// ROLL migration prototype. Compile and verify in TIA V19 before commissioning.
// No absolute M aliases: byte/word reads below preserve S5 overlapping memory.
TYPE "ROLL_TimerState"
VERSION : 0.1
STRUCT
    RemainingMs : LReal;
    BaseMs : Int;
    Mode : Int;
    Previous : Bool;
    Q : Bool;
END_STRUCT;
END_TYPE

TYPE "ROLL_CounterState"
VERSION : 0.1
STRUCT
    Value : Int;
    SetPrevious : Bool;
    UpPrevious : Bool;
    DownPrevious : Bool;
END_STRUCT;
END_TYPE

DATA_BLOCK "ROLL_State"
{ S7_Optimized_Access := 'TRUE' }
VERSION : 0.1
NON_RETAIN
VAR
    M : Array[0..255, 0..7] of Bool;
    S5Timers : Array[0..127] of "ROLL_TimerState";
    S5Counters : Array[0..127] of "ROLL_CounterState";
    CurrentProgram : Int := 1;
END_VAR
BEGIN
    M[0, 4] := TRUE;
END_DATA_BLOCK

DATA_BLOCK "ROLL_IO"
{ S7_Optimized_Access := 'TRUE' }
VERSION : 0.1
NON_RETAIN
VAR
    Input : Array[0..127, 0..7] of Bool;
    Output : Array[0..127, 0..7] of Bool;
    Simulation : Bool := TRUE;
    PhysicalOutputsEnabled : Bool := FALSE;
    PhysicalIoConfigured : Bool := FALSE;
    ConversionFault : Bool;
    FirstCycle : Bool := TRUE;
    RuntimeMemory : LReal;
    ClockMs : LReal;
    HmiElapsedMs : LReal;
    HmiLastHeartbeat : DInt;
END_VAR
BEGIN
END_DATA_BLOCK

// Flat, symbolic WinCC interface; TP900 control binding is a separate build step.
DATA_BLOCK "ROLL_HMI"
{ S7_Optimized_Access := 'TRUE' }
VERSION : 0.1
NON_RETAIN
VAR
    Heartbeat : DInt;
    Connected : Bool;
    ManualFunction : Int := 255;
    GroundHeld : Bool;
    WorkHeld : Bool;
    KeyF : Array[1..16] of Bool;
    SelectedProgram : Int := 1;
    RecipeCommand : Int := 1;
    RecipeRequest : DInt;
    RecipeAck : DInt;
    RecipeError : Int;
    CurrentProgram : Int := 1;
    ParameterRequest : DInt;
    ParameterAck : DInt;
    ParameterDb : Int := 15;
    ParameterIndex : Int;
    ParameterValue : DInt;
    ParameterCurrentValue : DInt;
    ParameterSlotPresent : Bool;
    ParameterError : Int;
    Dwell1Seconds : Int := 360;
    Drain1Seconds : Int := 90;
    Ultrasound1 : Bool := TRUE;
    Dwell2Seconds : Int := 240;
    Drain2Seconds : Int := 60;
    Dwell3Seconds : Int := 300;
    Drain3Seconds : Int := 120;
    Dry4Seconds : Int := 400;
    BasketMotion : Int := 1;
    BathLift : Bool;
    ProcessTimer1Units : Int;
    ProcessTimer2Units : Int;
    StatusM : Array[0..255, 0..7] of Bool;
    LogicalOutputs : Array[16..25, 0..7] of Bool;
END_VAR
BEGIN
END_DATA_BLOCK


DATA_BLOCK "ROLL_DB15"
{ S7_Optimized_Access := 'TRUE' }
VERSION : 0.1
NON_RETAIN
VAR
    DW : Array[0..131] of Word;
END_VAR
BEGIN
    DW[0] := W#16#FFFF;
    DW[1] := W#16#FFFF;
    DW[2] := W#16#FFFF;
    DW[3] := W#16#FFFF;
    DW[4] := W#16#FFFF;
    DW[5] := W#16#FFFF;
    DW[6] := W#16#FFFF;
    DW[7] := W#16#FFFF;
    DW[8] := W#16#FFFF;
    DW[9] := W#16#FFFF;
    DW[10] := W#16#FFFF;
    DW[11] := W#16#FFFF;
    DW[12] := W#16#FFFF;
    DW[13] := W#16#FFFF;
    DW[14] := W#16#FFFF;
    DW[15] := W#16#FFFF;
    DW[16] := W#16#FFFF;
    DW[17] := W#16#3360;
    DW[18] := W#16#FFFF;
    DW[19] := W#16#FFFF;
    DW[20] := W#16#FFFF;
    DW[21] := W#16#FFFF;
    DW[22] := W#16#FFFF;
    DW[23] := W#16#FFFF;
    DW[24] := W#16#1010;
    DW[25] := W#16#1020;
    DW[26] := W#16#FFFF;
    DW[27] := W#16#FFFF;
    DW[28] := W#16#FFFF;
    DW[29] := W#16#FFFF;
    DW[30] := W#16#FFFF;
    DW[31] := W#16#3120;
    DW[32] := W#16#3120;
    DW[33] := W#16#2900;
    DW[34] := W#16#FFFF;
    DW[35] := W#16#FFFF;
    DW[36] := W#16#FFFF;
    DW[37] := W#16#FFFF;
    DW[38] := W#16#FFFF;
    DW[39] := W#16#FFFF;
    DW[40] := W#16#FFFF;
    DW[41] := W#16#FFFF;
    DW[42] := W#16#FFFF;
    DW[43] := W#16#FFFF;
    DW[44] := W#16#FFFF;
    DW[45] := W#16#FFFF;
    DW[46] := W#16#FFFF;
    DW[47] := W#16#FFFF;
    DW[48] := W#16#FFFF;
    DW[49] := W#16#FFFF;
    DW[50] := W#16#FFFF;
    DW[51] := W#16#FFFF;
    DW[52] := W#16#FFFF;
    DW[53] := W#16#2120;
    DW[54] := W#16#2120;
    DW[55] := W#16#1010;
    DW[56] := W#16#2060;
    DW[57] := W#16#FFFF;
    DW[58] := W#16#3180;
    DW[59] := W#16#3180;
    DW[60] := W#16#2060;
    DW[61] := W#16#2600;
    DW[62] := W#16#2600;
    DW[63] := W#16#2010;
    DW[64] := W#16#FFFF;
    DW[65] := W#16#2015;
    DW[66] := W#16#FFFF;
    DW[67] := W#16#1050;
    DW[68] := W#16#FFFF;
    DW[69] := W#16#FFFF;
    DW[70] := W#16#FFFF;
    DW[71] := W#16#FFFF;
    DW[72] := W#16#FFFF;
    DW[73] := W#16#FFFF;
    DW[74] := W#16#FFFF;
    DW[75] := W#16#2600;
    DW[76] := W#16#FFFF;
    DW[77] := W#16#2300;
    DW[78] := W#16#FFFF;
    DW[79] := W#16#FFFF;
    DW[80] := W#16#FFFF;
    DW[81] := W#16#FFFF;
    DW[82] := W#16#FFFF;
    DW[83] := W#16#FFFF;
    DW[84] := W#16#FFFF;
    DW[85] := W#16#2120;
    DW[86] := W#16#FFFF;
    DW[87] := W#16#FFFF;
    DW[88] := W#16#FFFF;
    DW[89] := W#16#FFFF;
    DW[90] := W#16#FFFF;
    DW[91] := W#16#FFFF;
    DW[92] := W#16#FFFF;
    DW[93] := W#16#FFFF;
    DW[94] := W#16#FFFF;
    DW[95] := W#16#FFFF;
    DW[96] := W#16#FFFF;
    DW[97] := W#16#FFFF;
    DW[98] := W#16#FFFF;
    DW[99] := W#16#FFFF;
    DW[100] := W#16#FFFF;
    DW[101] := W#16#FFFF;
    DW[102] := W#16#2300;
    DW[103] := W#16#2300;
    DW[104] := W#16#FFFF;
    DW[105] := W#16#FFFF;
    DW[106] := W#16#2010;
    DW[107] := W#16#2015;
    DW[108] := W#16#FFFF;
    DW[109] := W#16#FFFF;
    DW[110] := W#16#FFFF;
    DW[111] := W#16#FFFF;
    DW[112] := W#16#FFFF;
    DW[113] := W#16#FFFF;
    DW[114] := W#16#FFFF;
    DW[115] := W#16#1050;
    DW[116] := W#16#1050;
    DW[117] := W#16#1050;
    DW[118] := W#16#FFFF;
    DW[119] := W#16#FFFF;
    DW[120] := W#16#FFFF;
    DW[121] := W#16#FFFF;
    DW[122] := W#16#FFFF;
    DW[123] := W#16#FFFF;
    DW[124] := W#16#FFFF;
    DW[125] := W#16#FFFF;
    DW[126] := W#16#FFFF;
    DW[127] := W#16#0038;
    DW[128] := W#16#0011;
    DW[129] := W#16#0011;
    DW[130] := W#16#3360;
    DW[131] := W#16#0000;
END_DATA_BLOCK

DATA_BLOCK "ROLL_DB19"
{ S7_Optimized_Access := 'TRUE' }
VERSION : 0.1
NON_RETAIN
VAR
    DW : Array[0..131] of Word;
END_VAR
BEGIN
    DW[0] := W#16#FFFF;
    DW[1] := W#16#0020;
    DW[2] := W#16#0014;
    DW[3] := W#16#FFFF;
    DW[4] := W#16#FFFF;
    DW[5] := W#16#FFFF;
    DW[6] := W#16#FFFF;
    DW[7] := W#16#FFFF;
    DW[8] := W#16#FFFF;
    DW[9] := W#16#FFFF;
    DW[10] := W#16#FFFF;
    DW[11] := W#16#FFFF;
    DW[12] := W#16#FFFF;
    DW[13] := W#16#FFFF;
    DW[14] := W#16#FFFF;
    DW[15] := W#16#FFFF;
    DW[16] := W#16#FFFF;
    DW[17] := W#16#FFFF;
    DW[18] := W#16#FFFF;
    DW[19] := W#16#FFFF;
    DW[20] := W#16#FFFF;
    DW[21] := W#16#FFFF;
    DW[22] := W#16#FFFF;
    DW[23] := W#16#FFFF;
    DW[24] := W#16#FFFF;
    DW[25] := W#16#FFFF;
    DW[26] := W#16#FFFF;
    DW[27] := W#16#FFFF;
    DW[28] := W#16#FFFF;
    DW[29] := W#16#FFFF;
    DW[30] := W#16#FFFF;
    DW[31] := W#16#FFFF;
    DW[32] := W#16#FFFF;
    DW[33] := W#16#FFFF;
    DW[34] := W#16#FFFF;
    DW[35] := W#16#FFFF;
    DW[36] := W#16#FFFF;
    DW[37] := W#16#FFFF;
    DW[38] := W#16#FFFF;
    DW[39] := W#16#FFFF;
    DW[40] := W#16#FFFF;
    DW[41] := W#16#FFFF;
    DW[42] := W#16#FFFF;
    DW[43] := W#16#FFFF;
    DW[44] := W#16#FFFF;
    DW[45] := W#16#FFFF;
    DW[46] := W#16#FFFF;
    DW[47] := W#16#FFFF;
    DW[48] := W#16#FFFF;
    DW[49] := W#16#FFFF;
    DW[50] := W#16#FFFF;
    DW[51] := W#16#FFFF;
    DW[52] := W#16#FFFF;
    DW[53] := W#16#FFFF;
    DW[54] := W#16#FFFF;
    DW[55] := W#16#FFFF;
    DW[56] := W#16#FFFF;
    DW[57] := W#16#FFFF;
    DW[58] := W#16#FFFF;
    DW[59] := W#16#FFFF;
    DW[60] := W#16#FFFF;
    DW[61] := W#16#FFFF;
    DW[62] := W#16#FFFF;
    DW[63] := W#16#FFFF;
    DW[64] := W#16#FFFF;
    DW[65] := W#16#FFFF;
    DW[66] := W#16#FFFF;
    DW[67] := W#16#FFFF;
    DW[68] := W#16#FFFF;
    DW[69] := W#16#FFFF;
    DW[70] := W#16#FFFF;
    DW[71] := W#16#FFFF;
    DW[72] := W#16#FFFF;
    DW[73] := W#16#FFFF;
    DW[74] := W#16#FFFF;
    DW[75] := W#16#FFFF;
    DW[76] := W#16#FFFF;
    DW[77] := W#16#FFFF;
    DW[78] := W#16#FFFF;
    DW[79] := W#16#FFFF;
    DW[80] := W#16#FFFF;
    DW[81] := W#16#FFFF;
    DW[82] := W#16#FFFF;
    DW[83] := W#16#FFFF;
    DW[84] := W#16#FFFF;
    DW[85] := W#16#FFFF;
    DW[86] := W#16#FFFF;
    DW[87] := W#16#FFFF;
    DW[88] := W#16#FFFF;
    DW[89] := W#16#FFFF;
    DW[90] := W#16#FFFF;
    DW[91] := W#16#FFFF;
    DW[92] := W#16#FFFF;
    DW[93] := W#16#FFFF;
    DW[94] := W#16#FFFF;
    DW[95] := W#16#FFFF;
    DW[96] := W#16#FFFF;
    DW[97] := W#16#FFFF;
    DW[98] := W#16#FFFF;
    DW[99] := W#16#FFFF;
    DW[100] := W#16#FFFF;
    DW[101] := W#16#FFFF;
    DW[102] := W#16#FFFF;
    DW[103] := W#16#FFFF;
    DW[104] := W#16#FFFF;
    DW[105] := W#16#FFFF;
    DW[106] := W#16#FFFF;
    DW[107] := W#16#FFFF;
    DW[108] := W#16#FFFF;
    DW[109] := W#16#FFFF;
    DW[110] := W#16#FFFF;
    DW[111] := W#16#FFFF;
    DW[112] := W#16#FFFF;
    DW[113] := W#16#FFFF;
    DW[114] := W#16#FFFF;
    DW[115] := W#16#FFFF;
    DW[116] := W#16#FFFF;
    DW[117] := W#16#FFFF;
    DW[118] := W#16#FFFF;
    DW[119] := W#16#FFFF;
    DW[120] := W#16#FFFF;
    DW[121] := W#16#FFFF;
    DW[122] := W#16#FFFF;
    DW[123] := W#16#FFFF;
    DW[124] := W#16#FFFF;
    DW[125] := W#16#FFFF;
    DW[126] := W#16#FFFF;
    DW[127] := W#16#FFFF;
    DW[128] := W#16#0001;
    DW[129] := W#16#0001;
    DW[130] := W#16#0020;
    DW[131] := W#16#0000;
END_DATA_BLOCK

DATA_BLOCK "ROLL_Recipe1"
{ S7_Optimized_Access := 'TRUE' }
VERSION : 0.1
NON_RETAIN
VAR
    DW : Array[0..41] of Word;
END_VAR
BEGIN
    DW[5] := W#16#2360;
    DW[9] := W#16#2090;
    DW[13] := W#16#0001;
    DW[17] := W#16#2240;
    DW[21] := W#16#2060;
    DW[25] := W#16#2300;
    DW[29] := W#16#2120;
    DW[33] := W#16#2400;
    DW[37] := W#16#0001;
    DW[41] := W#16#0000;
END_DATA_BLOCK

DATA_BLOCK "ROLL_Recipe2"
{ S7_Optimized_Access := 'TRUE' }
VERSION : 0.1
NON_RETAIN
VAR
    DW : Array[0..41] of Word;
END_VAR
BEGIN
    DW[5] := W#16#2360;
    DW[9] := W#16#2090;
    DW[13] := W#16#0001;
    DW[17] := W#16#2240;
    DW[21] := W#16#2060;
    DW[25] := W#16#2300;
    DW[29] := W#16#2120;
    DW[33] := W#16#2400;
    DW[37] := W#16#0001;
    DW[41] := W#16#0000;
END_DATA_BLOCK

DATA_BLOCK "ROLL_DB205"
{ S7_Optimized_Access := 'TRUE' }
VERSION : 0.1
NON_RETAIN
VAR
    DW : Array[0..41] of Word;
END_VAR
BEGIN
    DW[5] := W#16#2360;
    DW[9] := W#16#2090;
    DW[13] := W#16#0001;
    DW[17] := W#16#2240;
    DW[21] := W#16#2060;
    DW[25] := W#16#2300;
    DW[29] := W#16#2120;
    DW[33] := W#16#2400;
    DW[37] := W#16#0001;
    DW[41] := W#16#0000;
END_DATA_BLOCK

FUNCTION "ROLL_GetM" : Word
{ S7_Optimized_Access := 'TRUE' }
VERSION : 0.1
VAR_INPUT
    FirstByte : Int;
    Width : Int;
END_VAR
VAR_TEMP
    b : Int;
    n : Int;
    bit : Int;
    mask : Word;
    result : Word;
END_VAR
BEGIN
    #result := W#16#0000;
    IF (#FirstByte < 0) OR (#FirstByte > 255) OR ((#Width <> 8) AND (#Width <> 16)) OR ((#Width = 16) AND (#FirstByte > 254)) THEN
        "ROLL_IO".ConversionFault := TRUE;
        #ROLL_GetM := #result;
        RETURN;
    END_IF;
    FOR #n := 0 TO (#Width / 8) - 1 DO
        #b := #FirstByte + #n;
        FOR #bit := 0 TO 7 DO
            #mask := SHL(IN := W#16#0001, N := INT_TO_USINT(#bit + (#Width - 8 - 8 * #n)));
            IF "ROLL_State".M[#b, #bit] THEN #result := #result OR #mask; END_IF;
        END_FOR;
    END_FOR;
    #ROLL_GetM := #result;
END_FUNCTION

FUNCTION "ROLL_SetMWord" : Void
{ S7_Optimized_Access := 'TRUE' }
VERSION : 0.1
VAR_INPUT
    FirstByte : Int;
    Value : Word;
END_VAR
VAR_TEMP
    bit : Int;
END_VAR
BEGIN
    IF (#FirstByte < 0) OR (#FirstByte > 254) THEN
        "ROLL_IO".ConversionFault := TRUE;
        RETURN;
    END_IF;
    FOR #bit := 0 TO 7 DO
        "ROLL_State".M[#FirstByte, #bit] := (#Value AND SHL(IN := W#16#0001, N := INT_TO_USINT(#bit + 8))) <> W#16#0000;
        "ROLL_State".M[#FirstByte + 1, #bit] := (#Value AND SHL(IN := W#16#0001, N := INT_TO_USINT(#bit))) <> W#16#0000;
    END_FOR;
END_FUNCTION

FUNCTION "ROLL_GetDW" : Word
{ S7_Optimized_Access := 'TRUE' }
VERSION : 0.1
VAR_INPUT
    DbNumber : Int;
    Index : Int;
END_VAR
BEGIN
    #ROLL_GetDW := W#16#0000;
    IF (#Index < 0) OR (#Index > 131) THEN
        "ROLL_IO".ConversionFault := TRUE;
        RETURN;
    END_IF;
    CASE #DbNumber OF
        15: #ROLL_GetDW := "ROLL_DB15".DW[#Index];
        19: #ROLL_GetDW := "ROLL_DB19".DW[#Index];
        ELSE "ROLL_IO".ConversionFault := TRUE;
    END_CASE;
END_FUNCTION

FUNCTION "ROLL_DecodeBCD" : Int
{ S7_Optimized_Access := 'TRUE' }
VERSION : 0.1
VAR_INPUT
    Value : Word;
END_VAR
VAR_TEMP
    hundreds : Int;
    tens : Int;
    units : Int;
END_VAR
BEGIN
    #hundreds := WORD_TO_INT(SHR(IN := #Value AND W#16#0F00, N := 8));
    #tens := WORD_TO_INT(SHR(IN := #Value AND W#16#00F0, N := 4));
    #units := WORD_TO_INT(#Value AND W#16#000F);
    IF (#hundreds > 9) OR (#tens > 9) OR (#units > 9) THEN
        "ROLL_IO".ConversionFault := TRUE;
        #ROLL_DecodeBCD := -1;
    ELSE
        #ROLL_DecodeBCD := #hundreds * 100 + #tens * 10 + #units;
    END_IF;
END_FUNCTION

FUNCTION "ROLL_EncodeSeconds" : Word
{ S7_Optimized_Access := 'TRUE' }
VERSION : 0.1
VAR_INPUT
    Seconds : Int;
END_VAR
BEGIN
    IF (#Seconds < 0) OR (#Seconds > 999) THEN
        #ROLL_EncodeSeconds := W#16#FFFF;
    ELSE
        #ROLL_EncodeSeconds := W#16#2000 OR SHL(IN := INT_TO_WORD(#Seconds / 100), N := 8)
            OR SHL(IN := INT_TO_WORD((#Seconds / 10) MOD 10), N := 4) OR INT_TO_WORD(#Seconds MOD 10);
    END_IF;
END_FUNCTION

FUNCTION "ROLL_TimerOp" : Void
{ S7_Optimized_Access := 'TRUE' }
VERSION : 0.1
VAR_INPUT
    Number : Int;
    Operation : Int; // 0=SE on-delay; 1=SA off-delay; 2=R reset
    Signal : Bool;
    Preset : Word;
END_VAR
VAR_TEMP
    base : Int;
    count : Int;
    trigger : Bool;
END_VAR
BEGIN
    IF (#Number < 0) OR (#Number > 127) THEN
        "ROLL_IO".ConversionFault := TRUE;
        RETURN;
    END_IF;
    IF #Operation = 2 THEN
        IF #Signal THEN
            "ROLL_State".S5Timers[#Number].RemainingMs := 0.0;
            "ROLL_State".S5Timers[#Number].Q := FALSE;
        END_IF;
        RETURN;
    END_IF;
    #trigger := ((#Operation = 0) AND #Signal AND NOT "ROLL_State".S5Timers[#Number].Previous)
        OR ((#Operation = 1) AND NOT #Signal AND "ROLL_State".S5Timers[#Number].Previous);
    IF #trigger THEN
        #count := "ROLL_DecodeBCD"(Value := #Preset);
        #base := WORD_TO_INT(SHR(IN := #Preset AND W#16#F000, N := 12));
        CASE #base OF
            0: #base := 10;
            1: #base := 100;
            2: #base := 1000;
            3: #base := 10000;
            ELSE #base := 0;
        END_CASE;
        IF (#base = 0) OR (#count < 0) THEN
            "ROLL_IO".ConversionFault := TRUE;
            "ROLL_State".S5Timers[#Number].RemainingMs := 0.0;
            "ROLL_State".S5Timers[#Number].Q := FALSE;
            RETURN;
        END_IF;
        "ROLL_State".S5Timers[#Number].BaseMs := #base;
        "ROLL_State".S5Timers[#Number].RemainingMs := INT_TO_LREAL(#count) * INT_TO_LREAL(#base);
    END_IF;
    "ROLL_State".S5Timers[#Number].Mode := #Operation;
    IF #Operation = 0 THEN
        IF NOT #Signal THEN "ROLL_State".S5Timers[#Number].RemainingMs := 0.0; END_IF;
        "ROLL_State".S5Timers[#Number].Q := #Signal AND ("ROLL_State".S5Timers[#Number].RemainingMs <= 0.0);
    ELSIF #Operation = 1 THEN
        IF #Signal THEN "ROLL_State".S5Timers[#Number].RemainingMs := 0.0; END_IF;
        "ROLL_State".S5Timers[#Number].Q := #Signal OR ("ROLL_State".S5Timers[#Number].RemainingMs > 0.0);
    ELSE
        "ROLL_IO".ConversionFault := TRUE;
    END_IF;
    "ROLL_State".S5Timers[#Number].Previous := #Signal;
END_FUNCTION

FUNCTION "ROLL_TimerValue" : Word
{ S7_Optimized_Access := 'TRUE' }
VERSION : 0.1
VAR_INPUT
    Number : Int;
END_VAR
VAR_TEMP
    count : DInt;
END_VAR
BEGIN
    #ROLL_TimerValue := W#16#0000;
    IF (#Number < 0) OR (#Number > 127) THEN
        "ROLL_IO".ConversionFault := TRUE;
        RETURN;
    END_IF;
    IF "ROLL_State".S5Timers[#Number].BaseMs > 0 THEN
        #count := CEIL("ROLL_State".S5Timers[#Number].RemainingMs / INT_TO_LREAL("ROLL_State".S5Timers[#Number].BaseMs));
        #ROLL_TimerValue := DINT_TO_WORD(#count);
    END_IF;
END_FUNCTION

FUNCTION "ROLL_CounterOp" : Void
{ S7_Optimized_Access := 'TRUE' }
VERSION : 0.1
VAR_INPUT
    Number : Int;
    Operation : Int; // 0=S set; 1=R reset; 2=ZV up; 3=ZR down
    Signal : Bool;
    Preset : Word;
END_VAR
VAR_TEMP
    count : Int;
END_VAR
BEGIN
    IF (#Number < 0) OR (#Number > 127) THEN
        "ROLL_IO".ConversionFault := TRUE;
        RETURN;
    END_IF;
    CASE #Operation OF
        0:
            IF #Signal AND NOT "ROLL_State".S5Counters[#Number].SetPrevious THEN
                #count := "ROLL_DecodeBCD"(Value := #Preset);
                IF #count >= 0 THEN "ROLL_State".S5Counters[#Number].Value := #count; END_IF;
            END_IF;
            "ROLL_State".S5Counters[#Number].SetPrevious := #Signal;
        1:
            IF #Signal THEN "ROLL_State".S5Counters[#Number].Value := 0; END_IF;
        2:
            IF #Signal AND NOT "ROLL_State".S5Counters[#Number].UpPrevious AND ("ROLL_State".S5Counters[#Number].Value < 999) THEN
                "ROLL_State".S5Counters[#Number].Value := "ROLL_State".S5Counters[#Number].Value + 1;
            END_IF;
            "ROLL_State".S5Counters[#Number].UpPrevious := #Signal;
        3:
            IF #Signal AND NOT "ROLL_State".S5Counters[#Number].DownPrevious AND ("ROLL_State".S5Counters[#Number].Value > 0) THEN
                "ROLL_State".S5Counters[#Number].Value := "ROLL_State".S5Counters[#Number].Value - 1;
            END_IF;
            "ROLL_State".S5Counters[#Number].DownPrevious := #Signal;
        ELSE "ROLL_IO".ConversionFault := TRUE;
    END_CASE;
END_FUNCTION

FUNCTION "ROLL_AdvanceTime" : Void
{ S7_Optimized_Access := 'TRUE' }
VERSION : 0.1
VAR_INPUT
    DeltaMs : LReal;
END_VAR
VAR_TEMP
    n : Int;
END_VAR
BEGIN
    IF #DeltaMs < 0.0 THEN "ROLL_IO".ConversionFault := TRUE; RETURN; END_IF;
    FOR #n := 0 TO 127 DO
        IF "ROLL_State".S5Timers[#n].RemainingMs > 0.0 THEN
            "ROLL_State".S5Timers[#n].RemainingMs := "ROLL_State".S5Timers[#n].RemainingMs - #DeltaMs;
            IF "ROLL_State".S5Timers[#n].RemainingMs <= 0.0 THEN
                "ROLL_State".S5Timers[#n].RemainingMs := 0.0;
                "ROLL_State".S5Timers[#n].Q := "ROLL_State".S5Timers[#n].Mode = 0;
            END_IF;
        END_IF;
    END_FOR;
    "ROLL_IO".ClockMs := "ROLL_IO".ClockMs + #DeltaMs;
    WHILE "ROLL_IO".ClockMs >= 250.0 DO
        "ROLL_IO".ClockMs := "ROLL_IO".ClockMs - 250.0;
        "ROLL_State".M[3, 4] := NOT "ROLL_State".M[3, 4];
        IF NOT "ROLL_State".M[3, 4] THEN
            "ROLL_State".M[3, 5] := NOT "ROLL_State".M[3, 5];
            IF NOT "ROLL_State".M[3, 5] THEN
                "ROLL_State".M[3, 6] := NOT "ROLL_State".M[3, 6];
                IF NOT "ROLL_State".M[3, 6] THEN
                    "ROLL_State".M[3, 7] := NOT "ROLL_State".M[3, 7];
                END_IF;
            END_IF;
        END_IF;
    END_WHILE;
END_FUNCTION

FUNCTION "ROLL_FB69" : Void
{ S7_Optimized_Access := 'TRUE' }
VERSION : 0.1
BEGIN
    IF "ROLL_State".M[240, 0] AND "ROLL_State".M[240, 1] THEN
        "ROLL_SetMWord"(FirstByte := 240, Value := W#16#2005);
    ELSE
        "ROLL_SetMWord"(FirstByte := 240, Value := W#16#1005);
    END_IF;
END_FUNCTION

FUNCTION "ROLL_ShowRecipe" : Void
{ S7_Optimized_Access := 'TRUE' }
VERSION : 0.1
BEGIN
    "ROLL_HMI".CurrentProgram := "ROLL_State".CurrentProgram;
    "ROLL_HMI".SelectedProgram := "ROLL_State".CurrentProgram;
    "ROLL_HMI".Dwell1Seconds := "ROLL_DecodeBCD"(Value := "ROLL_DB205".DW[5]);
    "ROLL_HMI".Drain1Seconds := "ROLL_DecodeBCD"(Value := "ROLL_DB205".DW[9]);
    "ROLL_HMI".Dwell2Seconds := "ROLL_DecodeBCD"(Value := "ROLL_DB205".DW[17]);
    "ROLL_HMI".Drain2Seconds := "ROLL_DecodeBCD"(Value := "ROLL_DB205".DW[21]);
    "ROLL_HMI".Dwell3Seconds := "ROLL_DecodeBCD"(Value := "ROLL_DB205".DW[25]);
    "ROLL_HMI".Drain3Seconds := "ROLL_DecodeBCD"(Value := "ROLL_DB205".DW[29]);
    "ROLL_HMI".Dry4Seconds := "ROLL_DecodeBCD"(Value := "ROLL_DB205".DW[33]);
    "ROLL_HMI".Ultrasound1 := "ROLL_DB205".DW[13] = W#16#0001;
    "ROLL_HMI".BasketMotion := WORD_TO_INT("ROLL_DB205".DW[37]);
    "ROLL_HMI".BathLift := "ROLL_DB205".DW[41] = W#16#0001;
END_FUNCTION

FUNCTION "ROLL_FB90" : Void
{ S7_Optimized_Access := 'TRUE' }
VERSION : 0.1
BEGIN
    "ROLL_State".M[110, 0] := ("ROLL_DB205".DW[5] AND W#16#0FFF) <> W#16#0000;
    "ROLL_State".M[110, 1] := ("ROLL_DB205".DW[17] AND W#16#0FFF) <> W#16#0000;
    "ROLL_State".M[110, 2] := ("ROLL_DB205".DW[25] AND W#16#0FFF) <> W#16#0000;
    "ROLL_State".M[110, 3] := ("ROLL_DB205".DW[33] AND W#16#0FFF) <> W#16#0000;
    "ROLL_State".M[111, 0] := "ROLL_DB205".DW[37] = W#16#0001;
    "ROLL_State".M[111, 1] := "ROLL_DB205".DW[37] = W#16#0002;
    "ROLL_State".M[111, 2] := "ROLL_DB205".DW[37] = W#16#0003;
    "ROLL_State".M[111, 5] := "ROLL_DB205".DW[37] = W#16#0004;
    "ROLL_State".M[111, 3] := "ROLL_DB205".DW[41] = W#16#0001;
    "ROLL_State".M[111, 4] := "ROLL_DB205".DW[13] = W#16#0001;
    "ROLL_SetMWord"(FirstByte := 250, Value := W#16#0000);
END_FUNCTION

FUNCTION "ROLL_FB111" : Void
{ S7_Optimized_Access := 'TRUE' }
VERSION : 0.1
VAR_TEMP
    preset : Word;
    signal : Bool;
END_VAR
BEGIN
    #preset := W#16#2010;
    IF "ROLL_State".M[40, 5] THEN #preset := "ROLL_DB205".DW[5];
    ELSIF "ROLL_State".M[42, 1] THEN #preset := "ROLL_DB205".DW[17];
    ELSIF "ROLL_State".M[43, 5] THEN #preset := "ROLL_DB205".DW[25];
    ELSIF "ROLL_State".M[45, 2] THEN #preset := "ROLL_DB205".DW[33];
    END_IF;
    #signal := "ROLL_State".M[40, 5] OR "ROLL_State".M[42, 1] OR "ROLL_State".M[43, 5] OR "ROLL_State".M[45, 2]
        OR "ROLL_State".M[46, 5] OR "ROLL_State".M[48, 1] OR "ROLL_State".M[49, 5] OR "ROLL_State".M[51, 1];
    "ROLL_TimerOp"(Number := 1, Operation := 0, Signal := #signal, Preset := #preset);
    IF (WORD_TO_INT("ROLL_TimerValue"(Number := 1)) <= 7)
        AND ("ROLL_State".M[40, 5] OR "ROLL_State".M[42, 1] OR "ROLL_State".M[43, 5]) AND "ROLL_State".M[111, 5] THEN
        "ROLL_State".M[58, 5] := TRUE;
    END_IF;
    IF "ROLL_State".M[63, 1] AND "ROLL_IO".Input[13, 3] THEN "ROLL_State".M[58, 5] := FALSE; END_IF;
    #preset := W#16#2010;
    IF "ROLL_State".M[41, 1] THEN #preset := "ROLL_DB205".DW[9];
    ELSIF "ROLL_State".M[42, 5] THEN #preset := "ROLL_DB205".DW[21];
    ELSIF "ROLL_State".M[44, 1] THEN #preset := "ROLL_DB205".DW[29];
    END_IF;
    #signal := "ROLL_State".M[41, 1] OR "ROLL_State".M[42, 5] OR "ROLL_State".M[44, 1]
        OR "ROLL_State".M[45, 6] OR "ROLL_State".M[47, 1] OR "ROLL_State".M[48, 5] OR "ROLL_State".M[50, 1];
    "ROLL_TimerOp"(Number := 2, Operation := 0, Signal := #signal, Preset := #preset);
END_FUNCTION

FUNCTION "ROLL_PB2" : Void
{ S7_Optimized_Access := 'TRUE' }
VERSION : 0.1
VAR_TEMP
    r : Bool;
    a1 : Word;
    a2 : Word;
    activeDataBlock : Int;
    comparisonResults : Array[0..0] of Bool;
END_VAR
BEGIN
    #r := FALSE;
    #a1 := W#16#0000;
    #a2 := W#16#0000;
    #activeDataBlock := 0;
    // PB2, STEP 5 network 1
    #r := ((NOT "ROLL_State".M[0, 1]) AND "ROLL_State".S5Timers[11].Q);
    "ROLL_State".M[4, 1] := #r;
    // PB2, STEP 5 network 2
    #r := ((NOT "ROLL_State".M[4, 1]) OR "ROLL_IO".Input[1, 0]);
    "ROLL_State".M[3, 1] := #r;
    // PB2, STEP 5 network 3
    #r := ((((NOT "ROLL_State".M[31, 4]) AND "ROLL_IO".Input[0, 4] AND "ROLL_State".M[4, 1]) OR "ROLL_State".M[31, 5]) AND "ROLL_IO".Input[0, 2]);
    "ROLL_State".M[4, 4] := #r;
    // PB2, STEP 5 network 4
    #r := (NOT "ROLL_IO".Input[11, 7]);
    IF #r THEN "ROLL_State".M[5, 0] := TRUE; END_IF;
    #r := "ROLL_State".M[3, 1];
    IF #r THEN "ROLL_State".M[5, 0] := FALSE; END_IF;
    // PB2, STEP 5 network 5
    #r := (NOT "ROLL_IO".Input[13, 5]);
    IF #r THEN "ROLL_State".M[5, 1] := TRUE; END_IF;
    #r := "ROLL_State".M[3, 1];
    IF #r THEN "ROLL_State".M[5, 1] := FALSE; END_IF;
    // PB2, STEP 5 network 6
    #r := (NOT "ROLL_IO".Input[13, 0]);
    IF #r THEN "ROLL_State".M[5, 2] := TRUE; END_IF;
    #r := "ROLL_State".M[3, 1];
    IF #r THEN "ROLL_State".M[5, 2] := FALSE; END_IF;
    // PB2, STEP 5 network 7
    #r := (NOT "ROLL_IO".Input[8, 5]);
    IF #r THEN "ROLL_State".M[5, 3] := TRUE; END_IF;
    #r := "ROLL_State".M[3, 1];
    IF #r THEN "ROLL_State".M[5, 3] := FALSE; END_IF;
    // PB2, STEP 5 network 8
    #r := "ROLL_State".M[0, 3];
    IF #r THEN "ROLL_State".M[5, 4] := TRUE; END_IF;
    #r := "ROLL_State".M[3, 1];
    IF #r THEN "ROLL_State".M[5, 4] := FALSE; END_IF;
    // PB2, STEP 5 network 9
    #r := "ROLL_State".M[0, 3];
    IF #r THEN "ROLL_State".M[5, 5] := TRUE; END_IF;
    #r := "ROLL_State".M[3, 1];
    IF #r THEN "ROLL_State".M[5, 5] := FALSE; END_IF;
    // PB2, STEP 5 network 10
    #r := "ROLL_IO".Input[3, 6];
    IF #r THEN "ROLL_State".M[5, 6] := TRUE; END_IF;
    #r := "ROLL_State".M[3, 1];
    IF #r THEN "ROLL_State".M[5, 6] := FALSE; END_IF;
    // PB2, STEP 5 network 11
    #r := (NOT "ROLL_IO".Input[3, 7]);
    IF #r THEN "ROLL_State".M[5, 7] := TRUE; END_IF;
    #r := "ROLL_State".M[3, 1];
    IF #r THEN "ROLL_State".M[5, 7] := FALSE; END_IF;
    // PB2, STEP 5 network 12
    #r := (NOT "ROLL_IO".Input[5, 2]);
    IF #r THEN "ROLL_State".M[6, 0] := TRUE; END_IF;
    #r := ("ROLL_IO".Input[5, 2] AND "ROLL_State".M[3, 1]);
    IF #r THEN "ROLL_State".M[6, 0] := FALSE; END_IF;
    // PB2, STEP 5 network 13
    #r := ((NOT "ROLL_IO".Input[5, 3]) AND "ROLL_State".S5Timers[31].Q);
    IF #r THEN "ROLL_State".M[6, 1] := TRUE; END_IF;
    #r := "ROLL_State".M[3, 1];
    IF #r THEN "ROLL_State".M[6, 1] := FALSE; END_IF;
    // PB2, STEP 5 network 14
    #r := (NOT "ROLL_IO".Input[5, 4]);
    IF #r THEN "ROLL_State".M[6, 2] := TRUE; END_IF;
    #r := ("ROLL_IO".Input[5, 4] AND "ROLL_State".M[3, 1]);
    IF #r THEN "ROLL_State".M[6, 2] := FALSE; END_IF;
    // PB2, STEP 5 network 15
    #r := ((NOT "ROLL_IO".Input[5, 5]) AND "ROLL_State".M[40, 5] AND "ROLL_State".S5Timers[17].Q);
    IF #r THEN "ROLL_State".M[6, 3] := TRUE; END_IF;
    #r := "ROLL_State".M[3, 1];
    IF #r THEN "ROLL_State".M[6, 3] := FALSE; END_IF;
    // PB2, STEP 5 network 16
    #r := ((NOT "ROLL_IO".Input[6, 0]) AND "ROLL_State".S5Timers[32].Q);
    IF #r THEN "ROLL_State".M[6, 4] := TRUE; END_IF;
    #r := "ROLL_State".M[3, 1];
    IF #r THEN "ROLL_State".M[6, 4] := FALSE; END_IF;
    // PB2, STEP 5 network 17
    #r := ((NOT "ROLL_IO".Input[6, 2]) AND "ROLL_State".S5Timers[33].Q);
    IF #r THEN "ROLL_State".M[6, 5] := TRUE; END_IF;
    #r := "ROLL_State".M[3, 1];
    IF #r THEN "ROLL_State".M[6, 5] := FALSE; END_IF;
    // PB2, STEP 5 network 18
    #r := "ROLL_State".M[0, 3];
    IF #r THEN "ROLL_State".M[6, 6] := TRUE; END_IF;
    #r := "ROLL_State".M[3, 1];
    IF #r THEN "ROLL_State".M[6, 6] := FALSE; END_IF;
    // PB2, STEP 5 network 19
    #r := ((NOT "ROLL_State".M[0, 3]) AND "ROLL_State".S5Timers[35].Q);
    IF #r THEN "ROLL_State".M[6, 7] := TRUE; END_IF;
    #r := "ROLL_State".M[3, 1];
    IF #r THEN "ROLL_State".M[6, 7] := FALSE; END_IF;
    // PB2, STEP 5 network 20
    #r := ((NOT "ROLL_State".M[0, 3]) AND "ROLL_State".S5Timers[36].Q);
    IF #r THEN "ROLL_State".M[7, 0] := TRUE; END_IF;
    #r := "ROLL_State".M[3, 1];
    IF #r THEN "ROLL_State".M[7, 0] := FALSE; END_IF;
    // PB2, STEP 5 network 21
    #r := ((NOT "ROLL_State".M[0, 3]) AND "ROLL_State".M[48, 1] AND "ROLL_State".S5Timers[37].Q);
    IF #r THEN "ROLL_State".M[7, 1] := TRUE; END_IF;
    #r := "ROLL_State".M[3, 1];
    IF #r THEN "ROLL_State".M[7, 1] := FALSE; END_IF;
    // PB2, STEP 5 network 22
    #r := ((NOT "ROLL_State".M[0, 3]) AND "ROLL_State".S5Timers[38].Q);
    IF #r THEN "ROLL_State".M[7, 2] := TRUE; END_IF;
    #r := "ROLL_State".M[3, 1];
    IF #r THEN "ROLL_State".M[7, 2] := FALSE; END_IF;
    // PB2, STEP 5 network 23
    #r := ((NOT "ROLL_IO".Input[5, 6]) AND "ROLL_State".S5Timers[16].Q);
    IF #r THEN "ROLL_State".M[7, 3] := TRUE; END_IF;
    #r := ("ROLL_IO".Input[5, 6] AND "ROLL_State".M[3, 1]);
    IF #r THEN "ROLL_State".M[7, 3] := FALSE; END_IF;
    // PB2, STEP 5 network 24
    #r := "ROLL_State".M[0, 3];
    IF #r THEN "ROLL_State".M[7, 4] := TRUE; END_IF;
    #r := "ROLL_State".M[3, 1];
    IF #r THEN "ROLL_State".M[7, 4] := FALSE; END_IF;
    // PB2, STEP 5 network 25
    #r := "ROLL_State".M[0, 3];
    IF #r THEN "ROLL_State".M[7, 5] := TRUE; END_IF;
    #r := "ROLL_State".M[3, 1];
    IF #r THEN "ROLL_State".M[7, 5] := FALSE; END_IF;
    // PB2, STEP 5 network 26
    #r := "ROLL_State".M[0, 3];
    IF #r THEN "ROLL_State".M[7, 6] := TRUE; END_IF;
    #r := "ROLL_State".M[3, 1];
    IF #r THEN "ROLL_State".M[7, 6] := FALSE; END_IF;
    // PB2, STEP 5 network 27
    #r := (NOT "ROLL_IO".Input[6, 7]);
    IF #r THEN "ROLL_State".M[7, 7] := TRUE; END_IF;
    #r := "ROLL_State".M[3, 1];
    IF #r THEN "ROLL_State".M[7, 7] := FALSE; END_IF;
    // PB2, STEP 5 network 28
    #a2 := #a1;
    #a1 := W#16#1050;
    #r := ((NOT "ROLL_IO".Input[7, 6]) AND "ROLL_IO".Output[20, 5]);
    "ROLL_TimerOp"(Number := 30, Operation := 0, Signal := #r, Preset := #a1);
    #r := "ROLL_State".S5Timers[30].Q;
    IF #r THEN "ROLL_State".M[8, 6] := TRUE; END_IF;
    #r := "ROLL_State".M[3, 1];
    IF #r THEN "ROLL_State".M[8, 6] := FALSE; END_IF;
    // PB2, STEP 5 network 29
    #r := "ROLL_State".M[0, 3];
    IF #r THEN "ROLL_State".M[8, 7] := TRUE; END_IF;
    #r := "ROLL_State".M[3, 1];
    IF #r THEN "ROLL_State".M[8, 7] := FALSE; END_IF;
    // PB2, STEP 5 network 30
    #r := ((NOT "ROLL_IO".Input[13, 7]) AND "ROLL_State".M[4, 1]);
    IF #r THEN "ROLL_State".M[9, 0] := TRUE; END_IF;
    #r := ("ROLL_IO".Input[13, 7] AND "ROLL_State".M[3, 1]);
    IF #r THEN "ROLL_State".M[9, 0] := FALSE; END_IF;
    // PB2, STEP 5 network 31
    #r := "ROLL_State".M[0, 3];
    IF #r THEN "ROLL_State".M[9, 1] := TRUE; END_IF;
    #r := "ROLL_State".M[3, 1];
    IF #r THEN "ROLL_State".M[9, 1] := FALSE; END_IF;
    // PB2, STEP 5 network 32
    #r := ((NOT "ROLL_State".M[28, 4]) AND (NOT "ROLL_State".M[31, 5]) AND (((NOT "ROLL_State".M[20, 2]) AND ("ROLL_IO".Input[123, 5] OR "ROLL_IO".Input[123, 6])) OR "ROLL_State".M[70, 2] OR "ROLL_State".M[70, 3]) AND "ROLL_IO".Input[0, 4] AND "ROLL_State".M[4, 1]);
    IF #r THEN "ROLL_State".M[9, 2] := TRUE; END_IF;
    #r := "ROLL_State".M[3, 1];
    IF #r THEN "ROLL_State".M[9, 2] := FALSE; END_IF;
    // PB2, STEP 5 network 33
    #r := ("ROLL_State".M[4, 1] AND "ROLL_State".S5Timers[19].Q);
    IF #r THEN "ROLL_State".M[9, 3] := TRUE; END_IF;
    #r := "ROLL_State".M[3, 1];
    IF #r THEN "ROLL_State".M[9, 3] := FALSE; END_IF;
    // PB2, STEP 5 network 34
    #r := (((("ROLL_State".M[20, 4] OR "ROLL_State".M[20, 5]) AND "ROLL_IO".Input[0, 1] AND "ROLL_State".M[190, 6]) OR "ROLL_State".M[31, 5]) AND "ROLL_State".S5Timers[95].Q);
    "ROLL_State".M[9, 4] := #r;
    // PB2, STEP 5 network 35
    #r := "ROLL_State".M[0, 3];
    IF #r THEN "ROLL_State".M[9, 5] := TRUE; END_IF;
    #r := "ROLL_State".M[3, 1];
    IF #r THEN "ROLL_State".M[9, 5] := FALSE; END_IF;
    // PB2, STEP 5 network 36
    #r := "ROLL_State".M[0, 3];
    IF #r THEN "ROLL_State".M[9, 6] := TRUE; END_IF;
    #r := "ROLL_State".M[3, 1];
    IF #r THEN "ROLL_State".M[9, 6] := FALSE; END_IF;
    // PB2, STEP 5 network 37
    #r := "ROLL_State".M[0, 3];
    IF #r THEN "ROLL_State".M[9, 7] := TRUE; END_IF;
    #r := "ROLL_State".M[3, 1];
    IF #r THEN "ROLL_State".M[9, 7] := FALSE; END_IF;
    // PB2, STEP 5 network 38
    #r := ((NOT "ROLL_IO".Input[12, 0]) AND "ROLL_State".M[4, 1]);
    IF #r THEN "ROLL_State".M[10, 0] := TRUE; END_IF;
    #r := (((((NOT "ROLL_State".S5Timers[11].Q) AND "ROLL_IO".Input[3, 0]) OR "ROLL_IO".Input[12, 5]) AND "ROLL_State".M[3, 1]) OR (NOT "ROLL_State".M[4, 1]) OR "ROLL_State".M[0, 7]);
    IF #r THEN "ROLL_State".M[10, 0] := FALSE; END_IF;
    // PB2, STEP 5 network 39
    #r := ((NOT "ROLL_IO".Input[12, 6]) AND "ROLL_State".M[4, 1]);
    IF #r THEN "ROLL_State".M[10, 1] := TRUE; END_IF;
    #r := (((((NOT "ROLL_State".S5Timers[11].Q) AND "ROLL_IO".Input[3, 0]) OR "ROLL_IO".Input[12, 1]) AND "ROLL_State".M[3, 1]) OR (NOT "ROLL_State".M[4, 1]) OR "ROLL_State".M[0, 7]);
    IF #r THEN "ROLL_State".M[10, 1] := FALSE; END_IF;
    // PB2, STEP 5 network 40
    #r := "ROLL_State".M[0, 3];
    IF #r THEN "ROLL_State".M[10, 2] := TRUE; END_IF;
    #r := "ROLL_State".M[3, 1];
    IF #r THEN "ROLL_State".M[10, 2] := FALSE; END_IF;
    // PB2, STEP 5 network 41
    #r := "ROLL_State".M[0, 3];
    IF #r THEN "ROLL_State".M[10, 3] := TRUE; END_IF;
    #r := "ROLL_State".M[3, 1];
    IF #r THEN "ROLL_State".M[10, 3] := FALSE; END_IF;
    // PB2, STEP 5 network 42
    #r := "ROLL_State".M[0, 3];
    IF #r THEN "ROLL_State".M[10, 4] := TRUE; END_IF;
    #r := "ROLL_State".M[3, 1];
    IF #r THEN "ROLL_State".M[10, 4] := FALSE; END_IF;
    // PB2, STEP 5 network 43
    #r := "ROLL_State".M[0, 3];
    IF #r THEN "ROLL_State".M[10, 5] := TRUE; END_IF;
    #r := "ROLL_State".M[3, 1];
    IF #r THEN "ROLL_State".M[10, 5] := FALSE; END_IF;
    // PB2, STEP 5 network 44
    #r := "ROLL_State".M[0, 3];
    IF #r THEN "ROLL_State".M[10, 6] := TRUE; END_IF;
    #r := "ROLL_State".M[3, 1];
    IF #r THEN "ROLL_State".M[10, 6] := FALSE; END_IF;
    // PB2, STEP 5 network 45
    #r := "ROLL_State".M[0, 3];
    IF #r THEN "ROLL_State".M[10, 7] := TRUE; END_IF;
    #r := "ROLL_State".M[3, 1];
    IF #r THEN "ROLL_State".M[10, 7] := FALSE; END_IF;
    // PB2, STEP 5 network 46
    #r := ("ROLL_State".M[4, 1] AND "ROLL_State".M[63, 2]);
    IF #r THEN "ROLL_State".M[11, 0] := TRUE; END_IF;
    #r := "ROLL_State".M[3, 1];
    IF #r THEN "ROLL_State".M[11, 0] := FALSE; END_IF;
    // PB2, STEP 5 network 47
    #r := ("ROLL_IO".Input[13, 3] AND "ROLL_State".M[4, 1] AND "ROLL_State".S5Timers[112].Q);
    IF #r THEN "ROLL_State".M[11, 1] := TRUE; END_IF;
    #r := "ROLL_State".M[3, 1];
    IF #r THEN "ROLL_State".M[11, 1] := FALSE; END_IF;
    // PB2, STEP 5 network 48
    #r := ((NOT "ROLL_IO".Input[13, 3]) AND "ROLL_State".M[4, 1] AND "ROLL_State".S5Timers[15].Q);
    IF #r THEN "ROLL_State".M[11, 2] := TRUE; END_IF;
    #r := "ROLL_State".M[3, 1];
    IF #r THEN "ROLL_State".M[11, 2] := FALSE; END_IF;
    // PB2, STEP 5 network 49
    #r := ("ROLL_State".M[4, 1] AND "ROLL_State".M[63, 3]);
    IF #r THEN "ROLL_State".M[11, 3] := TRUE; END_IF;
    #r := "ROLL_State".M[3, 1];
    IF #r THEN "ROLL_State".M[11, 3] := FALSE; END_IF;
    // PB2, STEP 5 network 50
    #r := ("ROLL_State".M[190, 6] AND "ROLL_State".M[23, 2] AND "ROLL_State".M[60, 3]);
    IF #r THEN "ROLL_State".M[11, 4] := TRUE; END_IF;
    #r := "ROLL_State".M[3, 1];
    IF #r THEN "ROLL_State".M[11, 4] := FALSE; END_IF;
    // PB2, STEP 5 network 51
    #r := "ROLL_State".M[0, 3];
    IF #r THEN "ROLL_State".M[11, 5] := TRUE; END_IF;
    #r := "ROLL_State".M[3, 1];
    IF #r THEN "ROLL_State".M[11, 5] := FALSE; END_IF;
    // PB2, STEP 5 network 52
    #r := "ROLL_State".M[0, 3];
    IF #r THEN "ROLL_State".M[11, 6] := TRUE; END_IF;
    #r := "ROLL_State".M[3, 1];
    IF #r THEN "ROLL_State".M[11, 6] := FALSE; END_IF;
    // PB2, STEP 5 network 53
    #r := "ROLL_State".M[0, 3];
    IF #r THEN "ROLL_State".M[11, 7] := TRUE; END_IF;
    #r := "ROLL_State".M[3, 1];
    IF #r THEN "ROLL_State".M[11, 7] := FALSE; END_IF;
    // PB2, STEP 5 network 54
    #r := (NOT "ROLL_IO".Input[8, 3]);
    IF #r THEN "ROLL_State".M[12, 0] := TRUE; END_IF;
    #r := "ROLL_State".M[3, 1];
    IF #r THEN "ROLL_State".M[12, 0] := FALSE; END_IF;
    // PB2, STEP 5 network 55
    #r := ((NOT "ROLL_IO".Input[0, 7]) AND (NOT "ROLL_IO".Input[1, 4]) AND "ROLL_State".M[4, 4]);
    IF #r THEN "ROLL_State".M[12, 1] := TRUE; END_IF;
    #r := "ROLL_State".M[3, 1];
    IF #r THEN "ROLL_State".M[12, 1] := FALSE; END_IF;
    // PB2, STEP 5 network 56
    #r := "ROLL_State".M[0, 3];
    IF #r THEN "ROLL_State".M[12, 2] := TRUE; END_IF;
    #r := "ROLL_State".M[3, 1];
    IF #r THEN "ROLL_State".M[12, 2] := FALSE; END_IF;
    // PB2, STEP 5 network 57
    #r := "ROLL_State".M[0, 3];
    IF #r THEN "ROLL_State".M[12, 3] := TRUE; END_IF;
    #r := "ROLL_State".M[3, 1];
    IF #r THEN "ROLL_State".M[12, 3] := FALSE; END_IF;
    // PB2, STEP 5 network 58
    #r := "ROLL_State".M[0, 3];
    IF #r THEN "ROLL_State".M[13, 0] := TRUE; END_IF;
    #r := "ROLL_State".M[3, 1];
    IF #r THEN "ROLL_State".M[13, 0] := FALSE; END_IF;
    // PB2, STEP 5 network 59
    #r := (NOT "ROLL_IO".Input[3, 2]);
    IF #r THEN "ROLL_State".M[13, 1] := TRUE; END_IF;
    #r := "ROLL_State".M[3, 1];
    IF #r THEN "ROLL_State".M[13, 1] := FALSE; END_IF;
    // PB2, STEP 5 network 60
    #r := ((NOT "ROLL_IO".Input[4, 7]) AND "ROLL_IO".Input[0, 1] AND "ROLL_State".M[190, 6] AND "ROLL_State".M[27, 4]);
    IF #r THEN "ROLL_State".M[13, 2] := TRUE; END_IF;
    #r := "ROLL_State".M[3, 1];
    IF #r THEN "ROLL_State".M[13, 2] := FALSE; END_IF;
    // PB2, STEP 5 network 61
    #r := (NOT "ROLL_IO".Input[5, 0]);
    IF #r THEN "ROLL_State".M[13, 3] := TRUE; END_IF;
    #r := ("ROLL_IO".Input[5, 0] AND "ROLL_State".M[3, 1]);
    IF #r THEN "ROLL_State".M[13, 3] := FALSE; END_IF;
    // PB2, STEP 5 network 62
    #r := (NOT "ROLL_IO".Input[10, 7]);
    IF #r THEN "ROLL_State".M[13, 4] := TRUE; END_IF;
    #r := ("ROLL_IO".Input[10, 7] AND "ROLL_State".M[3, 1]);
    IF #r THEN "ROLL_State".M[13, 4] := FALSE; END_IF;
    // PB2, STEP 5 network 63
    #r := (NOT "ROLL_IO".Input[4, 5]);
    IF #r THEN "ROLL_State".M[13, 7] := TRUE; END_IF;
    #r := "ROLL_State".M[3, 1];
    IF #r THEN "ROLL_State".M[13, 7] := FALSE; END_IF;
    // PB2, STEP 5 network 64
    #a2 := #a1;
    #a1 := W#16#2020;
    #r := (((NOT "ROLL_IO".Input[10, 0]) OR (NOT "ROLL_IO".Input[10, 1]) OR (NOT "ROLL_IO".Input[10, 2]) OR (NOT "ROLL_IO".Input[10, 3])) AND "ROLL_IO".Output[19, 1]);
    "ROLL_TimerOp"(Number := 50, Operation := 0, Signal := #r, Preset := #a1);
    // PB2, STEP 5 network 65
    #r := ((NOT "ROLL_IO".Input[10, 0]) AND "ROLL_State".S5Timers[50].Q);
    IF #r THEN "ROLL_State".M[14, 0] := TRUE; END_IF;
    #r := "ROLL_State".M[3, 1];
    IF #r THEN "ROLL_State".M[14, 0] := FALSE; END_IF;
    // PB2, STEP 5 network 66
    #r := ((NOT "ROLL_IO".Input[10, 1]) AND "ROLL_State".S5Timers[50].Q);
    IF #r THEN "ROLL_State".M[14, 1] := TRUE; END_IF;
    #r := "ROLL_State".M[3, 1];
    IF #r THEN "ROLL_State".M[14, 1] := FALSE; END_IF;
    // PB2, STEP 5 network 67
    #r := ((NOT "ROLL_IO".Input[10, 2]) AND "ROLL_State".S5Timers[50].Q);
    IF #r THEN "ROLL_State".M[14, 2] := TRUE; END_IF;
    #r := "ROLL_State".M[3, 1];
    IF #r THEN "ROLL_State".M[14, 2] := FALSE; END_IF;
    // PB2, STEP 5 network 68
    #r := ((NOT "ROLL_IO".Input[10, 3]) AND "ROLL_State".S5Timers[50].Q);
    IF #r THEN "ROLL_State".M[14, 3] := TRUE; END_IF;
    #r := "ROLL_State".M[3, 1];
    IF #r THEN "ROLL_State".M[14, 3] := FALSE; END_IF;
    // PB2, STEP 5 network 69
    #r := "ROLL_State".M[0, 3];
    IF #r THEN "ROLL_State".M[15, 2] := TRUE; END_IF;
    #r := "ROLL_State".M[3, 1];
    IF #r THEN "ROLL_State".M[15, 2] := FALSE; END_IF;
    // PB2, STEP 5 network 70
    #r := "ROLL_State".M[0, 3];
    IF #r THEN "ROLL_State".M[15, 3] := TRUE; END_IF;
    #r := "ROLL_State".M[3, 1];
    IF #r THEN "ROLL_State".M[15, 3] := FALSE; END_IF;
    // PB2, STEP 5 network 71
    #r := "ROLL_State".M[0, 3];
    IF #r THEN "ROLL_State".M[15, 4] := TRUE; END_IF;
    #r := "ROLL_State".M[3, 1];
    IF #r THEN "ROLL_State".M[15, 4] := FALSE; END_IF;
    // PB2, STEP 5 network 72
    #r := (NOT "ROLL_IO".Input[4, 0]);
    IF #r THEN "ROLL_State".M[15, 5] := TRUE; END_IF;
    #r := "ROLL_State".M[3, 1];
    IF #r THEN "ROLL_State".M[15, 5] := FALSE; END_IF;
    // PB2, STEP 5 network 73
    #r := (NOT "ROLL_IO".Input[4, 1]);
    IF #r THEN "ROLL_State".M[15, 6] := TRUE; END_IF;
    #r := "ROLL_State".M[3, 1];
    IF #r THEN "ROLL_State".M[15, 6] := FALSE; END_IF;
    // PB2, STEP 5 network 74
    #r := (NOT "ROLL_IO".Input[4, 2]);
    IF #r THEN "ROLL_State".M[15, 7] := TRUE; END_IF;
    #r := "ROLL_State".M[3, 1];
    IF #r THEN "ROLL_State".M[15, 7] := FALSE; END_IF;
    // PB2, STEP 5 network 75
    #r := "ROLL_State".M[16, 0];
    IF #r THEN "ROLL_State".M[16, 0] := TRUE; END_IF;
    #r := "ROLL_State".M[3, 1];
    IF #r THEN "ROLL_State".M[16, 0] := FALSE; END_IF;
    // PB2, STEP 5 network 76
    #r := "ROLL_State".M[16, 1];
    IF #r THEN "ROLL_State".M[16, 1] := TRUE; END_IF;
    #r := "ROLL_State".M[3, 1];
    IF #r THEN "ROLL_State".M[16, 1] := FALSE; END_IF;
    // PB2, STEP 5 network 77
    #r := "ROLL_State".M[16, 2];
    IF #r THEN "ROLL_State".M[16, 2] := TRUE; END_IF;
    #r := "ROLL_State".M[3, 1];
    IF #r THEN "ROLL_State".M[16, 2] := FALSE; END_IF;
    // PB2, STEP 5 network 78
    #r := ("ROLL_State".M[34, 1] AND "ROLL_State".M[4, 1]);
    IF #r THEN "ROLL_State".M[16, 3] := TRUE; END_IF;
    #r := "ROLL_State".M[3, 1];
    IF #r THEN "ROLL_State".M[16, 3] := FALSE; END_IF;
    // PB2, STEP 5 network 79
    #r := "ROLL_State".M[16, 4];
    IF #r THEN "ROLL_State".M[16, 4] := TRUE; END_IF;
    #r := ((NOT "ROLL_IO".Input[123, 1]) AND (NOT "ROLL_IO".Input[123, 4]) AND (NOT "ROLL_IO".Input[123, 5]) AND (NOT "ROLL_IO".Input[123, 6]) AND (NOT "ROLL_IO".Input[125, 0]) AND (NOT "ROLL_IO".Input[125, 1]) AND "ROLL_State".M[3, 1]);
    IF #r THEN "ROLL_State".M[16, 4] := FALSE; END_IF;
    // PB2, STEP 5 network 80
    #r := "ROLL_State".M[16, 5];
    IF #r THEN "ROLL_State".M[16, 5] := TRUE; END_IF;
    #r := "ROLL_State".M[3, 1];
    IF #r THEN "ROLL_State".M[16, 5] := FALSE; END_IF;
    // PB2, STEP 5 network 81
    #r := ((NOT "ROLL_IO".Input[3, 4]) AND "ROLL_State".M[4, 1]);
    IF #r THEN "ROLL_State".M[16, 6] := TRUE; END_IF;
    #r := ("ROLL_IO".Input[3, 4] AND "ROLL_State".M[3, 1]);
    IF #r THEN "ROLL_State".M[16, 6] := FALSE; END_IF;
    // PB2, STEP 5 network 82
    #r := ((NOT "ROLL_IO".Input[3, 1]) AND ((("ROLL_State".M[190, 5] OR "ROLL_State".M[190, 6]) AND "ROLL_IO".Input[0, 1]) OR "ROLL_State".M[4, 4]) AND "ROLL_State".M[4, 1]);
    IF #r THEN "ROLL_State".M[16, 7] := TRUE; END_IF;
    #r := "ROLL_State".M[3, 1];
    IF #r THEN "ROLL_State".M[16, 7] := FALSE; END_IF;
    // PB2, STEP 5 network 83
    #r := ((NOT "ROLL_IO".Input[3, 5]) AND "ROLL_State".M[4, 1]);
    IF #r THEN "ROLL_State".M[17, 0] := TRUE; END_IF;
    #r := ("ROLL_IO".Input[3, 5] AND "ROLL_State".M[3, 1]);
    IF #r THEN "ROLL_State".M[17, 0] := FALSE; END_IF;
    // PB2, STEP 5 network 84
    #r := "ROLL_State".M[0, 3];
    IF #r THEN "ROLL_State".M[17, 1] := TRUE; END_IF;
    #r := "ROLL_State".M[3, 1];
    IF #r THEN "ROLL_State".M[17, 1] := FALSE; END_IF;
    // PB2, STEP 5 network 85
    #r := "ROLL_State".M[0, 3];
    IF #r THEN "ROLL_State".M[17, 2] := TRUE; END_IF;
    #r := "ROLL_State".M[3, 1];
    IF #r THEN "ROLL_State".M[17, 2] := FALSE; END_IF;
    // PB2, STEP 5 network 86
    #r := "ROLL_State".M[0, 3];
    IF #r THEN "ROLL_State".M[17, 3] := TRUE; END_IF;
    #r := "ROLL_State".M[3, 1];
    IF #r THEN "ROLL_State".M[17, 3] := FALSE; END_IF;
    // PB2, STEP 5 network 87
    #r := "ROLL_State".M[0, 3];
    IF #r THEN "ROLL_State".M[17, 4] := TRUE; END_IF;
    #r := "ROLL_State".M[3, 1];
    IF #r THEN "ROLL_State".M[17, 4] := FALSE; END_IF;
    // PB2, STEP 5 network 88
    #r := "ROLL_State".M[0, 3];
    IF #r THEN "ROLL_State".M[17, 5] := TRUE; END_IF;
    #r := "ROLL_State".M[3, 1];
    IF #r THEN "ROLL_State".M[17, 5] := FALSE; END_IF;
    // PB2, STEP 5 network 89
    #r := "ROLL_State".M[0, 3];
    IF #r THEN "ROLL_State".M[17, 6] := TRUE; END_IF;
    #r := "ROLL_State".M[3, 1];
    IF #r THEN "ROLL_State".M[17, 6] := FALSE; END_IF;
    // PB2, STEP 5 network 90
    #r := "ROLL_State".M[0, 3];
    IF #r THEN "ROLL_State".M[17, 7] := TRUE; END_IF;
    #r := "ROLL_State".M[3, 1];
    IF #r THEN "ROLL_State".M[17, 7] := FALSE; END_IF;
    // PB2, STEP 5 network 91
    #r := "ROLL_State".M[0, 3];
    IF #r THEN "ROLL_State".M[18, 0] := TRUE; END_IF;
    #r := "ROLL_State".M[3, 1];
    IF #r THEN "ROLL_State".M[18, 0] := FALSE; END_IF;
    // PB2, STEP 5 network 92
    #r := ((NOT "ROLL_IO".Input[14, 0]) AND ((("ROLL_State".M[190, 5] OR "ROLL_State".M[190, 6]) AND ("ROLL_State".M[23, 0] OR "ROLL_State".M[23, 1] OR "ROLL_State".M[23, 2] OR "ROLL_State".M[23, 3])) OR ("ROLL_State".M[16, 3] AND "ROLL_State".M[31, 4] AND "ROLL_State".M[37, 2]) OR "ROLL_State".M[74, 0]));
    IF #r THEN "ROLL_State".M[18, 1] := TRUE; END_IF;
    #r := "ROLL_State".M[3, 1];
    IF #r THEN "ROLL_State".M[18, 1] := FALSE; END_IF;
    // PB2, STEP 5 network 93
    #r := "ROLL_State".M[0, 3];
    IF #r THEN "ROLL_State".M[18, 2] := TRUE; END_IF;
    #r := "ROLL_State".M[3, 1];
    IF #r THEN "ROLL_State".M[18, 2] := FALSE; END_IF;
    // PB2, STEP 5 network 94
    #r := "ROLL_State".M[0, 3];
    IF #r THEN "ROLL_State".M[18, 3] := TRUE; END_IF;
    #r := "ROLL_State".M[3, 1];
    IF #r THEN "ROLL_State".M[18, 3] := FALSE; END_IF;
    // PB2, STEP 5 network 95
    #r := "ROLL_State".M[0, 3];
    IF #r THEN "ROLL_State".M[18, 4] := TRUE; END_IF;
    #r := "ROLL_State".M[3, 1];
    IF #r THEN "ROLL_State".M[18, 4] := FALSE; END_IF;
    // PB2, STEP 5 network 96
    #r := "ROLL_State".M[0, 3];
    IF #r THEN "ROLL_State".M[18, 5] := TRUE; END_IF;
    #r := "ROLL_State".M[3, 1];
    IF #r THEN "ROLL_State".M[18, 5] := FALSE; END_IF;
    // PB2, STEP 5 network 97
    #r := "ROLL_State".M[0, 3];
    IF #r THEN "ROLL_State".M[18, 6] := TRUE; END_IF;
    #r := "ROLL_State".M[3, 1];
    IF #r THEN "ROLL_State".M[18, 6] := FALSE; END_IF;
    // PB2, STEP 5 network 98
    #r := "ROLL_State".M[0, 3];
    IF #r THEN "ROLL_State".M[18, 7] := TRUE; END_IF;
    #r := "ROLL_State".M[3, 1];
    IF #r THEN "ROLL_State".M[18, 7] := FALSE; END_IF;
    // PB2, STEP 5 network 99
    #r := "ROLL_State".M[0, 3];
    IF #r THEN "ROLL_State".M[19, 0] := TRUE; END_IF;
    #r := "ROLL_State".M[3, 1];
    IF #r THEN "ROLL_State".M[19, 0] := FALSE; END_IF;
    // PB2, STEP 5 network 100
    #r := "ROLL_State".M[0, 3];
    IF #r THEN "ROLL_State".M[19, 1] := TRUE; END_IF;
    #r := "ROLL_State".M[3, 1];
    IF #r THEN "ROLL_State".M[19, 1] := FALSE; END_IF;
    // PB2, STEP 5 network 101
    #r := "ROLL_State".M[0, 3];
    IF #r THEN "ROLL_State".M[19, 2] := TRUE; END_IF;
    #r := "ROLL_State".M[3, 1];
    IF #r THEN "ROLL_State".M[19, 2] := FALSE; END_IF;
    // PB2, STEP 5 network 102
    #r := "ROLL_State".M[0, 3];
    IF #r THEN "ROLL_State".M[19, 3] := TRUE; END_IF;
    #r := "ROLL_State".M[3, 1];
    IF #r THEN "ROLL_State".M[19, 3] := FALSE; END_IF;
    // PB2, STEP 5 network 103
    #r := "ROLL_State".M[0, 3];
    IF #r THEN "ROLL_State".M[19, 4] := TRUE; END_IF;
    #r := "ROLL_State".M[3, 1];
    IF #r THEN "ROLL_State".M[19, 4] := FALSE; END_IF;
    // PB2, STEP 5 network 104
    #r := "ROLL_State".M[0, 3];
    IF #r THEN "ROLL_State".M[19, 5] := TRUE; END_IF;
    #r := "ROLL_State".M[3, 1];
    IF #r THEN "ROLL_State".M[19, 5] := FALSE; END_IF;
    // PB2, STEP 5 network 105
    #r := "ROLL_State".M[0, 3];
    IF #r THEN "ROLL_State".M[19, 6] := TRUE; END_IF;
    #r := "ROLL_State".M[3, 1];
    IF #r THEN "ROLL_State".M[19, 6] := FALSE; END_IF;
    // PB2, STEP 5 network 106
    #r := "ROLL_State".M[0, 3];
    IF #r THEN "ROLL_State".M[19, 7] := TRUE; END_IF;
    #r := "ROLL_State".M[3, 1];
    IF #r THEN "ROLL_State".M[19, 7] := FALSE; END_IF;
    // PB2, STEP 5 network 107
    RETURN;
END_FUNCTION

FUNCTION "ROLL_PB3" : Void
{ S7_Optimized_Access := 'TRUE' }
VERSION : 0.1
VAR_TEMP
    r : Bool;
    a1 : Word;
    a2 : Word;
    activeDataBlock : Int;
    comparisonResults : Array[0..15] of Bool;
END_VAR
BEGIN
    #r := FALSE;
    #a1 := W#16#0000;
    #a2 := W#16#0000;
    #activeDataBlock := 0;
    // PB3, STEP 5 network 1
    #a2 := #a1;
    #a1 := "ROLL_GetM"(FirstByte := 239, Width := 8);
    #a2 := #a1;
    #a1 := W#16#0001;
    #comparisonResults[0] := (WORD_TO_INT(#a2) = WORD_TO_INT(#a1));
    #r := #comparisonResults[0];
    "ROLL_State".M[20, 1] := #r;
    // PB3, STEP 5 network 2
    #a2 := #a1;
    #a1 := "ROLL_GetM"(FirstByte := 239, Width := 8);
    #a2 := #a1;
    #a1 := W#16#0002;
    #comparisonResults[1] := (WORD_TO_INT(#a2) = WORD_TO_INT(#a1));
    #r := #comparisonResults[1];
    "ROLL_State".M[20, 2] := #r;
    // PB3, STEP 5 network 3
    #a2 := #a1;
    #a1 := "ROLL_GetM"(FirstByte := 239, Width := 8);
    #a2 := #a1;
    #a1 := W#16#0003;
    #comparisonResults[2] := (WORD_TO_INT(#a2) = WORD_TO_INT(#a1));
    #r := #comparisonResults[2];
    "ROLL_State".M[20, 3] := #r;
    // PB3, STEP 5 network 4
    #a2 := #a1;
    #a1 := "ROLL_GetM"(FirstByte := 239, Width := 8);
    #a2 := #a1;
    #a1 := W#16#0004;
    #comparisonResults[3] := (WORD_TO_INT(#a2) = WORD_TO_INT(#a1));
    #r := #comparisonResults[3];
    "ROLL_State".M[20, 4] := #r;
    // PB3, STEP 5 network 5
    #a2 := #a1;
    #a1 := "ROLL_GetM"(FirstByte := 239, Width := 8);
    #a2 := #a1;
    #a1 := W#16#0005;
    #comparisonResults[4] := (WORD_TO_INT(#a2) = WORD_TO_INT(#a1));
    #r := #comparisonResults[4];
    "ROLL_State".M[20, 5] := #r;
    // PB3, STEP 5 network 6
    #a2 := #a1;
    #a1 := "ROLL_GetM"(FirstByte := 239, Width := 8);
    #a2 := #a1;
    #a1 := W#16#0007;
    #comparisonResults[5] := (WORD_TO_INT(#a2) = WORD_TO_INT(#a1));
    #r := #comparisonResults[5];
    "ROLL_State".M[20, 7] := #r;
    // PB3, STEP 5 network 7
    #a2 := #a1;
    #a1 := "ROLL_GetM"(FirstByte := 239, Width := 8);
    #a2 := #a1;
    #a1 := W#16#000A;
    #comparisonResults[6] := (WORD_TO_INT(#a2) = WORD_TO_INT(#a1));
    #r := #comparisonResults[6];
    "ROLL_State".M[22, 0] := #r;
    // PB3, STEP 5 network 8
    #a2 := #a1;
    #a1 := "ROLL_GetM"(FirstByte := 239, Width := 8);
    #a2 := #a1;
    #a1 := W#16#000B;
    #comparisonResults[7] := (WORD_TO_INT(#a2) = WORD_TO_INT(#a1));
    #r := #comparisonResults[7];
    "ROLL_State".M[22, 1] := #r;
    // PB3, STEP 5 network 9
    #a2 := #a1;
    #a1 := "ROLL_GetM"(FirstByte := 239, Width := 8);
    #a2 := #a1;
    #a1 := W#16#000C;
    #comparisonResults[8] := (WORD_TO_INT(#a2) = WORD_TO_INT(#a1));
    #r := #comparisonResults[8];
    "ROLL_State".M[22, 2] := #r;
    // PB3, STEP 5 network 10
    #a2 := #a1;
    #a1 := "ROLL_GetM"(FirstByte := 239, Width := 8);
    #a2 := #a1;
    #a1 := W#16#000D;
    #comparisonResults[9] := (WORD_TO_INT(#a2) = WORD_TO_INT(#a1));
    #r := #comparisonResults[9];
    "ROLL_State".M[22, 3] := #r;
    // PB3, STEP 5 network 11
    #a2 := #a1;
    #a1 := "ROLL_GetM"(FirstByte := 239, Width := 8);
    #a2 := #a1;
    #a1 := W#16#000E;
    #comparisonResults[10] := (WORD_TO_INT(#a2) = WORD_TO_INT(#a1));
    #r := #comparisonResults[10];
    "ROLL_State".M[22, 4] := #r;
    // PB3, STEP 5 network 12
    #a2 := #a1;
    #a1 := "ROLL_GetM"(FirstByte := 239, Width := 8);
    #a2 := #a1;
    #a1 := W#16#000F;
    #comparisonResults[11] := (WORD_TO_INT(#a2) = WORD_TO_INT(#a1));
    #r := #comparisonResults[11];
    "ROLL_State".M[22, 5] := #r;
    // PB3, STEP 5 network 13
    #a2 := #a1;
    #a1 := "ROLL_GetM"(FirstByte := 239, Width := 8);
    #a2 := #a1;
    #a1 := W#16#0014;
    #comparisonResults[12] := (WORD_TO_INT(#a2) = WORD_TO_INT(#a1));
    #r := #comparisonResults[12];
    "ROLL_State".M[23, 0] := #r;
    // PB3, STEP 5 network 14
    #a2 := #a1;
    #a1 := "ROLL_GetM"(FirstByte := 239, Width := 8);
    #a2 := #a1;
    #a1 := W#16#0015;
    #comparisonResults[13] := (WORD_TO_INT(#a2) = WORD_TO_INT(#a1));
    #r := #comparisonResults[13];
    "ROLL_State".M[23, 1] := #r;
    // PB3, STEP 5 network 15
    #a2 := #a1;
    #a1 := "ROLL_GetM"(FirstByte := 239, Width := 8);
    #a2 := #a1;
    #a1 := W#16#0016;
    #comparisonResults[14] := (WORD_TO_INT(#a2) = WORD_TO_INT(#a1));
    #r := #comparisonResults[14];
    "ROLL_State".M[23, 2] := #r;
    // PB3, STEP 5 network 16
    #a2 := #a1;
    #a1 := "ROLL_GetM"(FirstByte := 239, Width := 8);
    #a2 := #a1;
    #a1 := W#16#0017;
    #comparisonResults[15] := (WORD_TO_INT(#a2) = WORD_TO_INT(#a1));
    #r := #comparisonResults[15];
    "ROLL_State".M[23, 3] := #r;
    // PB3, STEP 5 network 17
    RETURN;
END_FUNCTION

FUNCTION "ROLL_PB4" : Void
{ S7_Optimized_Access := 'TRUE' }
VERSION : 0.1
VAR_TEMP
    r : Bool;
    a1 : Word;
    a2 : Word;
    activeDataBlock : Int;
    comparisonResults : Array[0..24] of Bool;
END_VAR
BEGIN
    #r := FALSE;
    #a1 := W#16#0000;
    #a2 := W#16#0000;
    #activeDataBlock := 0;
    // PB4, STEP 5 network 1
    #a2 := #a1;
    #a1 := "ROLL_GetM"(FirstByte := 239, Width := 8);
    #a2 := #a1;
    #a1 := W#16#001E;
    #comparisonResults[0] := (WORD_TO_INT(#a2) = WORD_TO_INT(#a1));
    #r := #comparisonResults[0];
    "ROLL_State".M[23, 5] := #r;
    // PB4, STEP 5 network 2
    #a2 := #a1;
    #a1 := "ROLL_GetM"(FirstByte := 239, Width := 8);
    #a2 := #a1;
    #a1 := W#16#001F;
    #comparisonResults[1] := (WORD_TO_INT(#a2) = WORD_TO_INT(#a1));
    #r := #comparisonResults[1];
    "ROLL_State".M[23, 6] := #r;
    // PB4, STEP 5 network 3
    #a2 := #a1;
    #a1 := "ROLL_GetM"(FirstByte := 239, Width := 8);
    #a2 := #a1;
    #a1 := W#16#0023;
    #comparisonResults[2] := (WORD_TO_INT(#a2) = WORD_TO_INT(#a1));
    #r := #comparisonResults[2];
    "ROLL_State".M[24, 0] := #r;
    // PB4, STEP 5 network 4
    #a2 := #a1;
    #a1 := "ROLL_GetM"(FirstByte := 239, Width := 8);
    #a2 := #a1;
    #a1 := W#16#0024;
    #comparisonResults[3] := (WORD_TO_INT(#a2) = WORD_TO_INT(#a1));
    #r := #comparisonResults[3];
    "ROLL_State".M[24, 1] := #r;
    // PB4, STEP 5 network 5
    #a2 := #a1;
    #a1 := "ROLL_GetM"(FirstByte := 239, Width := 8);
    #a2 := #a1;
    #a1 := W#16#0025;
    #comparisonResults[4] := (WORD_TO_INT(#a2) = WORD_TO_INT(#a1));
    #r := #comparisonResults[4];
    "ROLL_State".M[24, 2] := #r;
    // PB4, STEP 5 network 6
    #a2 := #a1;
    #a1 := "ROLL_GetM"(FirstByte := 239, Width := 8);
    #a2 := #a1;
    #a1 := W#16#0026;
    #comparisonResults[5] := (WORD_TO_INT(#a2) = WORD_TO_INT(#a1));
    #r := #comparisonResults[5];
    "ROLL_State".M[24, 3] := #r;
    // PB4, STEP 5 network 7
    #a2 := #a1;
    #a1 := "ROLL_GetM"(FirstByte := 239, Width := 8);
    #a2 := #a1;
    #a1 := W#16#0027;
    #comparisonResults[6] := (WORD_TO_INT(#a2) = WORD_TO_INT(#a1));
    #r := #comparisonResults[6];
    "ROLL_State".M[24, 4] := #r;
    // PB4, STEP 5 network 8
    #a2 := #a1;
    #a1 := "ROLL_GetM"(FirstByte := 239, Width := 8);
    #a2 := #a1;
    #a1 := W#16#0032;
    #comparisonResults[7] := (WORD_TO_INT(#a2) = WORD_TO_INT(#a1));
    #r := #comparisonResults[7];
    "ROLL_State".M[25, 0] := #r;
    // PB4, STEP 5 network 9
    #a2 := #a1;
    #a1 := "ROLL_GetM"(FirstByte := 239, Width := 8);
    #a2 := #a1;
    #a1 := W#16#0033;
    #comparisonResults[8] := (WORD_TO_INT(#a2) = WORD_TO_INT(#a1));
    #r := #comparisonResults[8];
    "ROLL_State".M[25, 1] := #r;
    // PB4, STEP 5 network 10
    #a2 := #a1;
    #a1 := "ROLL_GetM"(FirstByte := 239, Width := 8);
    #a2 := #a1;
    #a1 := W#16#0034;
    #comparisonResults[9] := (WORD_TO_INT(#a2) = WORD_TO_INT(#a1));
    #r := #comparisonResults[9];
    "ROLL_State".M[25, 2] := #r;
    // PB4, STEP 5 network 11
    #a2 := #a1;
    #a1 := "ROLL_GetM"(FirstByte := 239, Width := 8);
    #a2 := #a1;
    #a1 := W#16#0035;
    #comparisonResults[10] := (WORD_TO_INT(#a2) = WORD_TO_INT(#a1));
    #r := #comparisonResults[10];
    "ROLL_State".M[25, 3] := #r;
    // PB4, STEP 5 network 12
    #a2 := #a1;
    #a1 := "ROLL_GetM"(FirstByte := 239, Width := 8);
    #a2 := #a1;
    #a1 := W#16#0037;
    #comparisonResults[11] := (WORD_TO_INT(#a2) = WORD_TO_INT(#a1));
    #r := #comparisonResults[11];
    "ROLL_State".M[25, 4] := #r;
    // PB4, STEP 5 network 13
    #a2 := #a1;
    #a1 := "ROLL_GetM"(FirstByte := 239, Width := 8);
    #a2 := #a1;
    #a1 := W#16#0038;
    #comparisonResults[12] := (WORD_TO_INT(#a2) = WORD_TO_INT(#a1));
    #r := #comparisonResults[12];
    "ROLL_State".M[25, 5] := #r;
    // PB4, STEP 5 network 14
    #a2 := #a1;
    #a1 := "ROLL_GetM"(FirstByte := 239, Width := 8);
    #a2 := #a1;
    #a1 := W#16#0039;
    #comparisonResults[13] := (WORD_TO_INT(#a2) = WORD_TO_INT(#a1));
    #r := #comparisonResults[13];
    "ROLL_State".M[25, 6] := #r;
    // PB4, STEP 5 network 15
    #a2 := #a1;
    #a1 := "ROLL_GetM"(FirstByte := 239, Width := 8);
    #a2 := #a1;
    #a1 := W#16#003A;
    #comparisonResults[14] := (WORD_TO_INT(#a2) = WORD_TO_INT(#a1));
    #r := #comparisonResults[14];
    "ROLL_State".M[25, 7] := #r;
    // PB4, STEP 5 network 16
    #a2 := #a1;
    #a1 := "ROLL_GetM"(FirstByte := 239, Width := 8);
    #a2 := #a1;
    #a1 := W#16#003C;
    #comparisonResults[15] := (WORD_TO_INT(#a2) = WORD_TO_INT(#a1));
    #r := #comparisonResults[15];
    "ROLL_State".M[26, 0] := #r;
    // PB4, STEP 5 network 17
    #a2 := #a1;
    #a1 := "ROLL_GetM"(FirstByte := 239, Width := 8);
    #a2 := #a1;
    #a1 := W#16#003D;
    #comparisonResults[16] := (WORD_TO_INT(#a2) = WORD_TO_INT(#a1));
    #r := #comparisonResults[16];
    "ROLL_State".M[26, 1] := #r;
    // PB4, STEP 5 network 18
    #a2 := #a1;
    #a1 := "ROLL_GetM"(FirstByte := 239, Width := 8);
    #a2 := #a1;
    #a1 := W#16#003E;
    #comparisonResults[17] := (WORD_TO_INT(#a2) = WORD_TO_INT(#a1));
    #r := #comparisonResults[17];
    "ROLL_State".M[26, 2] := #r;
    // PB4, STEP 5 network 19
    #a2 := #a1;
    #a1 := "ROLL_GetM"(FirstByte := 239, Width := 8);
    #a2 := #a1;
    #a1 := W#16#003F;
    #comparisonResults[18] := (WORD_TO_INT(#a2) = WORD_TO_INT(#a1));
    #r := #comparisonResults[18];
    "ROLL_State".M[26, 3] := #r;
    // PB4, STEP 5 network 20
    #a2 := #a1;
    #a1 := "ROLL_GetM"(FirstByte := 239, Width := 8);
    #a2 := #a1;
    #a1 := W#16#0041;
    #comparisonResults[19] := (WORD_TO_INT(#a2) = WORD_TO_INT(#a1));
    #r := #comparisonResults[19];
    "ROLL_State".M[26, 5] := #r;
    // PB4, STEP 5 network 21
    #a2 := #a1;
    #a1 := "ROLL_GetM"(FirstByte := 239, Width := 8);
    #a2 := #a1;
    #a1 := W#16#0042;
    #comparisonResults[20] := (WORD_TO_INT(#a2) = WORD_TO_INT(#a1));
    #r := #comparisonResults[20];
    "ROLL_State".M[26, 6] := #r;
    // PB4, STEP 5 network 22
    #a2 := #a1;
    #a1 := "ROLL_GetM"(FirstByte := 239, Width := 8);
    #a2 := #a1;
    #a1 := W#16#0045;
    #comparisonResults[21] := (WORD_TO_INT(#a2) = WORD_TO_INT(#a1));
    #r := #comparisonResults[21];
    "ROLL_State".M[27, 1] := #r;
    // PB4, STEP 5 network 23
    #a2 := #a1;
    #a1 := "ROLL_GetM"(FirstByte := 239, Width := 8);
    #a2 := #a1;
    #a1 := W#16#0048;
    #comparisonResults[22] := (WORD_TO_INT(#a2) = WORD_TO_INT(#a1));
    #r := #comparisonResults[22];
    "ROLL_State".M[27, 4] := #r;
    // PB4, STEP 5 network 24
    #a2 := #a1;
    #a1 := "ROLL_GetM"(FirstByte := 239, Width := 8);
    #a2 := #a1;
    #a1 := W#16#0049;
    #comparisonResults[23] := (WORD_TO_INT(#a2) = WORD_TO_INT(#a1));
    #r := #comparisonResults[23];
    "ROLL_State".M[27, 5] := #r;
    // PB4, STEP 5 network 25
    #a2 := #a1;
    #a1 := "ROLL_GetM"(FirstByte := 239, Width := 8);
    #a2 := #a1;
    #a1 := W#16#0063;
    #comparisonResults[24] := (WORD_TO_INT(#a2) = WORD_TO_INT(#a1));
    #r := #comparisonResults[24];
    "ROLL_State".M[27, 7] := #r;
    // PB4, STEP 5 network 26
    RETURN;
END_FUNCTION

FUNCTION "ROLL_PB7" : Void
{ S7_Optimized_Access := 'TRUE' }
VERSION : 0.1
VAR_TEMP
    r : Bool;
    a1 : Word;
    a2 : Word;
    activeDataBlock : Int;
    comparisonResults : Array[0..0] of Bool;
END_VAR
BEGIN
    #r := FALSE;
    #a1 := W#16#0000;
    #a2 := W#16#0000;
    #activeDataBlock := 0;
    // PB7, STEP 5 network 1
    #r := ((NOT "ROLL_State".M[70, 2]) AND (NOT "ROLL_State".M[70, 3]) AND (NOT "ROLL_State".M[70, 4]) AND (NOT "ROLL_State".M[70, 6]) AND "ROLL_IO".Input[11, 0] AND "ROLL_IO".Input[11, 6] AND "ROLL_IO".Input[13, 3] AND "ROLL_State".M[63, 1]);
    "ROLL_State".M[28, 0] := #r;
    // PB7, STEP 5 network 2
    #r := ("ROLL_IO".Input[12, 1] AND "ROLL_IO".Input[12, 7]);
    "ROLL_State".M[28, 1] := #r;
    // PB7, STEP 5 network 3
    #r := ((NOT "ROLL_IO".Output[112, 5]) AND ((NOT "ROLL_IO".Output[112, 0]) OR (NOT "ROLL_State".M[31, 4])));
    "ROLL_State".M[28, 2] := #r;
    // PB7, STEP 5 network 4
    #r := (((NOT "ROLL_IO".Output[113, 0]) AND (NOT "ROLL_IO".Output[113, 1]) AND (NOT "ROLL_IO".Output[113, 3]) AND (NOT "ROLL_IO".Output[113, 5]) AND (NOT "ROLL_IO".Input[123, 5]) AND (NOT "ROLL_IO".Input[123, 6]) AND "ROLL_IO".Output[113, 2] AND "ROLL_IO".Output[113, 4] AND "ROLL_IO".Input[124, 1] AND "ROLL_IO".Input[124, 4]) OR "ROLL_State".M[0, 4]);
    "ROLL_State".M[240, 0] := #r;
    // PB7, STEP 5 network 5
    #r := ((((NOT "ROLL_IO".Output[113, 2]) AND "ROLL_IO".Output[113, 3] AND "ROLL_IO".Input[123, 5] AND "ROLL_IO".Input[124, 1] AND "ROLL_IO".Input[124, 4]) OR ((NOT "ROLL_IO".Output[113, 3]) AND "ROLL_IO".Output[113, 2] AND "ROLL_IO".Input[124, 1] AND "ROLL_IO".Input[124, 5]) OR "ROLL_State".M[0, 4]) AND "ROLL_State".M[20, 2]);
    "ROLL_State".M[240, 1] := #r;
    // PB7, STEP 5 network 6
    #r := ("ROLL_State".M[240, 0] OR "ROLL_State".M[240, 1]);
    "ROLL_State".M[28, 3] := #r;
    // PB7, STEP 5 network 7
    #r := ("ROLL_State".M[28, 0] AND "ROLL_State".M[28, 1] AND "ROLL_State".M[28, 2] AND "ROLL_State".M[28, 3]);
    "ROLL_State".M[28, 4] := #r;
    // PB7, STEP 5 network 8
    #r := ("ROLL_IO".Input[10, 7] AND "ROLL_IO".Input[3, 4] AND "ROLL_IO".Input[3, 5] AND "ROLL_IO".Input[3, 7]);
    "ROLL_State".M[28, 5] := #r;
    // PB7, STEP 5 network 9
    #r := ((NOT "ROLL_State".M[13, 4]) AND (NOT "ROLL_State".M[16, 6]) AND (NOT "ROLL_State".M[5, 7]) AND "ROLL_State".M[28, 5]);
    "ROLL_State".M[28, 6] := #r;
    // PB7, STEP 5 network 10
    #r := (("ROLL_IO".Input[0, 2] AND "ROLL_IO".Input[0, 4]) OR "ROLL_IO".Input[0, 1]);
    IF #r THEN "ROLL_State".M[29, 0] := TRUE; END_IF;
    #r := (NOT "ROLL_State".M[28, 6]);
    IF #r THEN "ROLL_State".M[29, 0] := FALSE; END_IF;
    // PB7, STEP 5 network 11
    #r := ("ROLL_State".M[29, 0] AND "ROLL_State".S5Timers[13].Q);
    "ROLL_State".M[29, 1] := #r;
    // PB7, STEP 5 network 12
    #r := (NOT "ROLL_State".M[12, 1]);
    "ROLL_State".M[30, 0] := #r;
    // PB7, STEP 5 network 13
    #r := "ROLL_State".M[0, 4];
    "ROLL_State".M[30, 1] := #r;
    // PB7, STEP 5 network 14
    #r := ((NOT "ROLL_State".M[6, 1]) AND (NOT "ROLL_State".M[6, 3]) AND (NOT "ROLL_State".M[6, 4]) AND (NOT "ROLL_State".M[6, 5]) AND (NOT "ROLL_State".M[6, 6]) AND (NOT "ROLL_State".M[6, 7]) AND (NOT "ROLL_State".M[7, 0]) AND (NOT "ROLL_State".M[7, 1]) AND (NOT "ROLL_State".M[7, 2]) AND (NOT "ROLL_State".M[7, 3]) AND (NOT "ROLL_State".M[7, 7]));
    "ROLL_State".M[30, 2] := #r;
    // PB7, STEP 5 network 15
    #r := ((NOT "ROLL_IO".Input[3, 6]) AND (NOT "ROLL_State".M[5, 6]));
    "ROLL_State".M[30, 3] := #r;
    // PB7, STEP 5 network 16
    #r := (("ROLL_State".M[30, 0] AND "ROLL_State".M[30, 1] AND "ROLL_State".M[30, 2] AND "ROLL_State".M[30, 3]) OR "ROLL_IO".Input[0, 0] OR "ROLL_IO".Input[0, 6]);
    "ROLL_State".M[30, 5] := #r;
    // PB7, STEP 5 network 17
    #r := ((NOT "ROLL_State".M[11, 0]) AND (NOT "ROLL_State".M[13, 1]) AND (NOT "ROLL_State".M[13, 3]) AND (NOT "ROLL_State".M[5, 0]) AND (NOT "ROLL_State".M[5, 1]) AND (NOT "ROLL_State".M[5, 2]));
    "ROLL_State".M[30, 6] := #r;
    // PB7, STEP 5 network 18
    #r := ((NOT "ROLL_State".M[11, 1]) AND (NOT "ROLL_State".M[5, 3]) AND (NOT "ROLL_State".M[9, 1]) AND (NOT "ROLL_State".M[9, 2]) AND (NOT "ROLL_State".M[9, 3]) AND "ROLL_IO".Input[8, 5] AND "ROLL_State".M[28, 6]);
    "ROLL_State".M[30, 7] := #r;
    // PB7, STEP 5 network 19
    #r := ((NOT "ROLL_State".M[12, 0]) AND (NOT "ROLL_State".M[9, 0]));
    "ROLL_State".M[31, 0] := #r;
    // PB7, STEP 5 network 20
    #r := ((NOT "ROLL_State".M[87, 5]) AND (NOT "ROLL_State".M[88, 1]) AND (NOT "ROLL_State".M[88, 3]) AND (NOT "ROLL_State".M[88, 4]) AND (NOT "ROLL_State".M[88, 5]) AND (NOT "ROLL_State".M[88, 6]));
    "ROLL_State".M[31, 2] := #r;
    // PB7, STEP 5 network 21
    #r := ("ROLL_State".M[30, 5] AND "ROLL_State".M[30, 6] AND "ROLL_State".M[30, 7] AND "ROLL_State".M[31, 0] AND "ROLL_State".M[31, 2]);
    "ROLL_State".M[31, 1] := #r;
    // PB7, STEP 5 network 22
    #r := (("ROLL_State".M[28, 4] OR "ROLL_State".M[31, 5]) AND "ROLL_IO".Input[0, 4] AND "ROLL_State".M[4, 4]);
    IF #r THEN "ROLL_State".M[31, 4] := TRUE; END_IF;
    #r := ((NOT "ROLL_IO".Input[0, 2]) OR (NOT "ROLL_IO".Input[0, 3]) OR (NOT "ROLL_State".M[29, 0]) OR (NOT "ROLL_State".M[31, 1]));
    IF #r THEN "ROLL_State".M[31, 4] := FALSE; END_IF;
    // PB7, STEP 5 network 23
    #r := "ROLL_State".M[31, 4];
    IF #r THEN "ROLL_State".M[31, 5] := TRUE; END_IF;
    #r := (((NOT "ROLL_State".M[31, 4]) AND (((NOT "ROLL_State".M[37, 2]) AND "ROLL_State".M[37, 1]) OR "ROLL_State".M[37, 0]) AND "ROLL_State".M[28, 4]) OR (NOT "ROLL_IO".Input[0, 2]));
    IF #r THEN "ROLL_State".M[31, 5] := FALSE; END_IF;
    // PB7, STEP 5 network 24
    #r := "ROLL_State".M[52, 3];
    IF #r THEN "ROLL_State".M[31, 6] := TRUE; END_IF;
    #r := ((NOT "ROLL_IO".Input[14, 0]) AND "ROLL_IO".Input[12, 1]);
    IF #r THEN "ROLL_State".M[31, 6] := FALSE; END_IF;
    // PB7, STEP 5 network 25
    #r := "ROLL_State".M[31, 5];
    "ROLL_IO".Output[16, 6] := #r;
    // PB7, STEP 5 network 26
    #r := "ROLL_State".M[40, 0];
    "ROLL_IO".Output[16, 7] := #r;
    // PB7, STEP 5 network 27
    RETURN;
END_FUNCTION

FUNCTION "ROLL_PB8" : Void
{ S7_Optimized_Access := 'TRUE' }
VERSION : 0.1
VAR_TEMP
    r : Bool;
    a1 : Word;
    a2 : Word;
    activeDataBlock : Int;
    comparisonResults : Array[0..0] of Bool;
END_VAR
BEGIN
    #r := FALSE;
    #a1 := W#16#0000;
    #a2 := W#16#0000;
    #activeDataBlock := 0;
    // PB8, STEP 5 network 1
    #r := ("ROLL_State".M[37, 7] OR "ROLL_State".M[38, 0] OR "ROLL_State".M[39, 7] OR "ROLL_State".M[40, 0] OR "ROLL_State".M[40, 1] OR "ROLL_State".M[40, 4] OR "ROLL_State".M[41, 0] OR "ROLL_State".M[41, 6] OR "ROLL_State".M[41, 7] OR "ROLL_State".M[42, 2] OR "ROLL_State".M[42, 3]);
    "ROLL_State".M[33, 0] := #r;
    // PB8, STEP 5 network 2
    #r := (((NOT "ROLL_State".M[16, 0]) AND (NOT "ROLL_State".M[16, 1]) AND (NOT "ROLL_State".M[16, 4]) AND "ROLL_State".M[37, 2]) OR "ROLL_State".M[37, 3] OR "ROLL_State".M[37, 5] OR "ROLL_State".M[37, 6] OR "ROLL_State".M[39, 4] OR "ROLL_State".M[39, 5] OR "ROLL_State".M[40, 2] OR "ROLL_State".M[40, 3] OR "ROLL_State".M[40, 6] OR "ROLL_State".M[40, 7] OR "ROLL_State".M[41, 2] OR "ROLL_State".M[42, 0] OR "ROLL_State".M[42, 4]);
    "ROLL_State".M[33, 1] := #r;
    // PB8, STEP 5 network 3
    #a2 := #a1;
    #a1 := W#16#2030;
    #r := ((NOT "ROLL_State".M[3, 1]) AND ("ROLL_State".M[33, 0] OR "ROLL_State".M[42, 6] OR "ROLL_State".M[43, 4] OR "ROLL_State".M[43, 6] OR "ROLL_State".M[43, 7] OR "ROLL_State".M[44, 2] OR "ROLL_State".M[45, 0] OR "ROLL_State".M[45, 1] OR "ROLL_State".M[45, 5] OR "ROLL_State".M[45, 7] OR "ROLL_State".M[46, 1] OR "ROLL_State".M[46, 4] OR "ROLL_State".M[46, 6] OR "ROLL_State".M[52, 1] OR "ROLL_State".M[52, 2] OR "ROLL_State".M[53, 3]) AND "ROLL_IO".Input[0, 2] AND "ROLL_State".M[29, 0]);
    "ROLL_TimerOp"(Number := 40, Operation := 0, Signal := #r, Preset := #a1);
    // PB8, STEP 5 network 4
    #a2 := #a1;
    #a1 := W#16#2030;
    #r := ((NOT "ROLL_State".M[3, 1]) AND (((NOT "ROLL_IO".Input[11, 2]) AND "ROLL_State".M[52, 0]) OR ((NOT "ROLL_State".M[15, 1]) AND "ROLL_State".M[53, 1]) OR "ROLL_State".M[33, 1] OR "ROLL_State".M[43, 0] OR "ROLL_State".M[43, 2] OR "ROLL_State".M[43, 3] OR "ROLL_State".M[44, 0] OR "ROLL_State".M[44, 7] OR "ROLL_State".M[45, 3] OR "ROLL_State".M[45, 4] OR "ROLL_State".M[46, 2] OR "ROLL_State".M[46, 3] OR "ROLL_State".M[46, 7] OR "ROLL_State".M[47, 3] OR "ROLL_State".M[52, 3] OR "ROLL_State".M[53, 2] OR "ROLL_State".M[53, 5] OR "ROLL_State".M[53, 6]) AND "ROLL_IO".Input[0, 2] AND "ROLL_State".M[29, 0]);
    "ROLL_TimerOp"(Number := 41, Operation := 0, Signal := #r, Preset := #a1);
    // PB8, STEP 5 network 5
    #r := ("ROLL_State".S5Timers[40].Q OR "ROLL_State".S5Timers[41].Q);
    IF #r THEN "ROLL_State".M[34, 1] := TRUE; END_IF;
    #r := ((NOT "ROLL_IO".Input[0, 2]) OR "ROLL_State".M[3, 1]);
    IF #r THEN "ROLL_State".M[34, 1] := FALSE; END_IF;
    // PB8, STEP 5 network 6
    RETURN;
END_FUNCTION

FUNCTION "ROLL_PB9" : Void
{ S7_Optimized_Access := 'TRUE' }
VERSION : 0.1
VAR_TEMP
    r : Bool;
    a1 : Word;
    a2 : Word;
    activeDataBlock : Int;
    comparisonResults : Array[0..0] of Bool;
END_VAR
BEGIN
    #r := FALSE;
    #a1 := W#16#0000;
    #a2 := W#16#0000;
    #activeDataBlock := 0;
    // PB9, STEP 5 network 1
    #r := ((NOT "ROLL_State".M[32, 1]) AND (NOT "ROLL_State".M[32, 2]) AND "ROLL_IO".Input[0, 2]);
    "ROLL_State".M[32, 0] := #r;
    // PB9, STEP 5 network 2
    #r := "ROLL_State".M[32, 0];
    IF #r THEN "ROLL_State".M[32, 1] := TRUE; END_IF;
    #r := ((NOT "ROLL_IO".Input[0, 2]) OR "ROLL_IO".Input[0, 1] OR "ROLL_State".M[32, 2]);
    IF #r THEN "ROLL_State".M[32, 1] := FALSE; END_IF;
    // PB9, STEP 5 network 3
    #r := ((NOT "ROLL_IO".Input[0, 2]) OR "ROLL_IO".Input[0, 1]);
    "ROLL_State".M[32, 2] := #r;
    // PB9, STEP 5 network 4
    #r := ((NOT "ROLL_State".M[12, 0]) AND (NOT "ROLL_State".M[5, 0]) AND (NOT "ROLL_State".M[5, 2]) AND (NOT "ROLL_State".M[9, 0]));
    "ROLL_State".M[35, 1] := #r;
    // PB9, STEP 5 network 5
    #r := "ROLL_IO".Input[0, 4];
    IF #r THEN "ROLL_State".M[35, 2] := TRUE; END_IF;
    #r := ((NOT "ROLL_State".M[29, 0]) OR (NOT "ROLL_State".M[31, 5]) OR (NOT "ROLL_State".M[35, 1]) OR "ROLL_State".M[16, 3]);
    IF #r THEN "ROLL_State".M[35, 2] := FALSE; END_IF;
    // PB9, STEP 5 network 6
    #r := ("ROLL_State".M[32, 0] OR "ROLL_State".M[53, 6]);
    IF #r THEN "ROLL_State".M[37, 0] := TRUE; END_IF;
    #r := ("ROLL_State".M[32, 2] OR "ROLL_State".M[37, 1] OR "ROLL_State".M[38, 0] OR "ROLL_State".M[39, 5]);
    IF #r THEN "ROLL_State".M[37, 0] := FALSE; END_IF;
    // PB9, STEP 5 network 7
    #r := ((NOT "ROLL_IO".Input[123, 5]) AND (NOT "ROLL_IO".Input[123, 6]) AND (NOT "ROLL_State".M[53, 6]) AND "ROLL_State".M[31, 5] AND "ROLL_State".M[35, 2] AND "ROLL_State".M[37, 0]);
    IF #r THEN "ROLL_State".M[37, 1] := TRUE; END_IF;
    #r := ("ROLL_State".M[32, 2] OR "ROLL_State".M[37, 2] OR "ROLL_State".M[39, 6]);
    IF #r THEN "ROLL_State".M[37, 1] := FALSE; END_IF;
    // PB9, STEP 5 network 8
    #r := ((NOT "ROLL_IO".Output[113, 3]) AND (NOT "ROLL_State".M[9, 1]) AND (("ROLL_IO".Input[0, 5] AND "ROLL_IO".Input[14, 3] AND "ROLL_State".M[0, 4]) OR ("ROLL_IO".Input[123, 4] AND "ROLL_IO".Input[124, 4] AND "ROLL_State".M[0, 3])) AND "ROLL_State".M[35, 2] AND "ROLL_State".M[37, 1]);
    IF #r THEN "ROLL_State".M[37, 2] := TRUE; END_IF;
    #r := ("ROLL_State".M[32, 2] OR "ROLL_State".M[37, 3]);
    IF #r THEN "ROLL_State".M[37, 2] := FALSE; END_IF;
    // PB9, STEP 5 network 9
    #r := ((NOT "ROLL_State".M[16, 0]) AND (NOT "ROLL_State".M[16, 1]) AND (NOT "ROLL_State".M[16, 4]) AND (NOT "ROLL_State".M[191, 5]) AND "ROLL_IO".Input[14, 0] AND "ROLL_State".M[190, 1] AND "ROLL_State".M[191, 4] AND "ROLL_State".M[35, 2] AND "ROLL_State".M[37, 2]);
    IF #r THEN "ROLL_State".M[37, 3] := TRUE; END_IF;
    #r := ("ROLL_State".M[32, 2] OR "ROLL_State".M[37, 5] OR "ROLL_State".M[40, 0]);
    IF #r THEN "ROLL_State".M[37, 3] := FALSE; END_IF;
    // PB9, STEP 5 network 10
    #r := ((NOT "ROLL_IO".Input[123, 5]) AND (NOT "ROLL_IO".Input[123, 6]) AND "ROLL_IO".Input[124, 1] AND "ROLL_IO".Input[124, 4] AND "ROLL_State".M[0, 3] AND "ROLL_State".M[35, 2] AND "ROLL_State".M[37, 3]);
    IF #r THEN "ROLL_State".M[37, 5] := TRUE; END_IF;
    #r := ("ROLL_State".M[32, 2] OR "ROLL_State".M[37, 6]);
    IF #r THEN "ROLL_State".M[37, 5] := FALSE; END_IF;
    // PB9, STEP 5 network 11
    #r := ((NOT "ROLL_IO".Output[113, 2]) AND "ROLL_IO".Output[113, 3] AND "ROLL_State".M[35, 2] AND "ROLL_State".M[37, 5] AND "ROLL_State".S5Timers[18].Q);
    IF #r THEN "ROLL_State".M[37, 6] := TRUE; END_IF;
    #r := ("ROLL_State".M[32, 2] OR "ROLL_State".M[37, 7]);
    IF #r THEN "ROLL_State".M[37, 6] := FALSE; END_IF;
    // PB9, STEP 5 network 12
    #r := ((NOT "ROLL_State".M[37, 5]) AND "ROLL_State".M[35, 2] AND "ROLL_State".M[37, 6]);
    IF #r THEN "ROLL_State".M[37, 7] := TRUE; END_IF;
    #r := ("ROLL_State".M[32, 2] OR "ROLL_State".M[38, 0]);
    IF #r THEN "ROLL_State".M[37, 7] := FALSE; END_IF;
    // PB9, STEP 5 network 13
    #r := ((NOT "ROLL_State".M[70, 2]) AND (((NOT "ROLL_IO".Output[113, 2]) AND "ROLL_IO".Output[113, 3] AND "ROLL_IO".Input[124, 4] AND "ROLL_State".M[28, 4] AND "ROLL_State".M[37, 0]) OR ("ROLL_State".M[37, 7] AND "ROLL_State".S5Timers[20].Q)) AND "ROLL_IO".Input[123, 5] AND "ROLL_State".M[35, 2]);
    IF #r THEN "ROLL_State".M[38, 0] := TRUE; END_IF;
    #r := ("ROLL_State".M[32, 2] OR "ROLL_State".M[39, 4]);
    IF #r THEN "ROLL_State".M[38, 0] := FALSE; END_IF;
    // PB9, STEP 5 network 14
    #r := ((NOT "ROLL_IO".Input[124, 5]) AND "ROLL_IO".Input[124, 4] AND "ROLL_State".M[35, 2] AND "ROLL_State".M[38, 0]);
    IF #r THEN "ROLL_State".M[39, 4] := TRUE; END_IF;
    #r := ("ROLL_State".M[32, 2] OR "ROLL_State".M[39, 5]);
    IF #r THEN "ROLL_State".M[39, 4] := FALSE; END_IF;
    // PB9, STEP 5 network 15
    #r := ((NOT "ROLL_IO".Input[124, 4]) AND (("ROLL_State".M[28, 4] AND "ROLL_State".M[37, 0]) OR "ROLL_State".M[39, 4]) AND "ROLL_IO".Input[124, 5] AND "ROLL_State".M[35, 2]);
    IF #r THEN "ROLL_State".M[39, 5] := TRUE; END_IF;
    #r := ("ROLL_State".M[32, 2] OR "ROLL_State".M[39, 6]);
    IF #r THEN "ROLL_State".M[39, 5] := FALSE; END_IF;
    // PB9, STEP 5 network 16
    #r := ((NOT "ROLL_IO".Input[124, 2]) AND "ROLL_IO".Input[11, 0] AND "ROLL_IO".Input[11, 6] AND "ROLL_IO".Input[12, 1] AND "ROLL_IO".Input[12, 7] AND "ROLL_IO".Input[124, 1] AND "ROLL_State".M[35, 2] AND "ROLL_State".M[39, 5]);
    IF #r THEN "ROLL_State".M[39, 6] := TRUE; END_IF;
    #r := ("ROLL_State".M[32, 2] OR "ROLL_State".M[39, 7]);
    IF #r THEN "ROLL_State".M[39, 6] := FALSE; END_IF;
    // PB9, STEP 5 network 17
    #r := ((NOT "ROLL_IO".Input[124, 1]) AND "ROLL_IO".Input[124, 2] AND "ROLL_State".M[35, 2] AND "ROLL_State".M[39, 6]);
    IF #r THEN "ROLL_State".M[39, 7] := TRUE; END_IF;
    #r := ("ROLL_State".M[32, 2] OR "ROLL_State".M[40, 0]);
    IF #r THEN "ROLL_State".M[39, 7] := FALSE; END_IF;
    // PB9, STEP 5 network 18
    #r := ((NOT "ROLL_IO".Input[12, 5]) AND ("ROLL_State".M[37, 3] OR "ROLL_State".M[39, 7]) AND "ROLL_IO".Input[11, 0] AND "ROLL_IO".Input[11, 6] AND "ROLL_IO".Input[12, 1] AND "ROLL_IO".Input[12, 7] AND "ROLL_State".M[35, 2]);
    IF #r THEN "ROLL_State".M[40, 0] := TRUE; END_IF;
    #r := ("ROLL_State".M[32, 2] OR "ROLL_State".M[40, 1]);
    IF #r THEN "ROLL_State".M[40, 0] := FALSE; END_IF;
    // PB9, STEP 5 network 19
    #r := ("ROLL_IO".Input[12, 5] AND "ROLL_IO".Input[12, 7] AND "ROLL_State".M[35, 2] AND "ROLL_State".M[40, 0]);
    IF #r THEN "ROLL_State".M[40, 1] := TRUE; END_IF;
    #r := ("ROLL_State".M[32, 2] OR "ROLL_State".M[40, 2] OR "ROLL_State".M[41, 6] OR "ROLL_State".M[43, 2] OR "ROLL_State".M[44, 7] OR "ROLL_State".M[46, 2] OR "ROLL_State".M[47, 6] OR "ROLL_State".M[49, 2] OR "ROLL_State".M[50, 6]);
    IF #r THEN "ROLL_State".M[40, 1] := FALSE; END_IF;
    // PB9, STEP 5 network 20
    #r := ((NOT "ROLL_IO".Input[11, 1]) AND "ROLL_IO".Input[11, 0] AND "ROLL_State".M[110, 0] AND "ROLL_State".M[35, 2] AND "ROLL_State".M[40, 1] AND "ROLL_State".M[63, 1]);
    IF #r THEN "ROLL_State".M[40, 2] := TRUE; END_IF;
    #r := ("ROLL_State".M[32, 2] OR "ROLL_State".M[40, 3]);
    IF #r THEN "ROLL_State".M[40, 2] := FALSE; END_IF;
    // PB9, STEP 5 network 21
    #r := ("ROLL_IO".Input[11, 1] AND "ROLL_IO".Input[11, 6] AND "ROLL_State".M[35, 2] AND "ROLL_State".M[40, 2]);
    IF #r THEN "ROLL_State".M[40, 3] := TRUE; END_IF;
    #r := ("ROLL_State".M[32, 2] OR "ROLL_State".M[40, 4]);
    IF #r THEN "ROLL_State".M[40, 3] := FALSE; END_IF;
    // PB9, STEP 5 network 22
    #r := ((NOT "ROLL_IO".Input[12, 1]) AND "ROLL_IO".Input[12, 5] AND "ROLL_State".M[35, 2] AND "ROLL_State".M[40, 3]);
    IF #r THEN "ROLL_State".M[40, 4] := TRUE; END_IF;
    #r := ("ROLL_State".M[32, 2] OR "ROLL_State".M[40, 5]);
    IF #r THEN "ROLL_State".M[40, 4] := FALSE; END_IF;
    // PB9, STEP 5 network 23
    #r := ("ROLL_IO".Input[12, 1] AND "ROLL_IO".Input[12, 7] AND "ROLL_State".M[35, 2] AND "ROLL_State".M[40, 4]);
    IF #r THEN "ROLL_State".M[40, 5] := TRUE; END_IF;
    #r := ("ROLL_State".M[32, 2] OR "ROLL_State".M[40, 6]);
    IF #r THEN "ROLL_State".M[40, 5] := FALSE; END_IF;
    // PB9, STEP 5 network 24
    #r := ("ROLL_State".M[35, 2] AND "ROLL_State".M[40, 5] AND "ROLL_State".S5Timers[1].Q);
    IF #r THEN "ROLL_State".M[40, 6] := TRUE; END_IF;
    #r := ("ROLL_State".M[32, 2] OR "ROLL_State".M[40, 7]);
    IF #r THEN "ROLL_State".M[40, 6] := FALSE; END_IF;
    // PB9, STEP 5 network 25
    #r := ("ROLL_State".M[35, 2] AND "ROLL_State".M[40, 6]);
    IF #r THEN "ROLL_State".M[40, 7] := TRUE; END_IF;
    #r := ("ROLL_State".M[32, 2] OR "ROLL_State".M[41, 0]);
    IF #r THEN "ROLL_State".M[40, 7] := FALSE; END_IF;
    // PB9, STEP 5 network 26
    #r := ((NOT "ROLL_IO".Input[12, 5]) AND (("ROLL_IO".Input[13, 3] AND "ROLL_State".M[63, 1]) OR (NOT "ROLL_State".M[111, 5])) AND "ROLL_State".M[35, 2] AND "ROLL_State".M[40, 7]);
    IF #r THEN "ROLL_State".M[41, 0] := TRUE; END_IF;
    #r := ("ROLL_State".M[32, 2] OR "ROLL_State".M[41, 1]);
    IF #r THEN "ROLL_State".M[41, 0] := FALSE; END_IF;
    // PB9, STEP 5 network 27
    #r := ("ROLL_IO".Input[12, 5] AND "ROLL_IO".Input[12, 7] AND "ROLL_State".M[35, 2] AND "ROLL_State".M[41, 0]);
    IF #r THEN "ROLL_State".M[41, 1] := TRUE; END_IF;
    #r := ("ROLL_State".M[32, 2] OR "ROLL_State".M[41, 2]);
    IF #r THEN "ROLL_State".M[41, 1] := FALSE; END_IF;
    // PB9, STEP 5 network 28
    #r := ("ROLL_State".M[35, 2] AND "ROLL_State".M[41, 1] AND "ROLL_State".S5Timers[2].Q);
    IF #r THEN "ROLL_State".M[41, 2] := TRUE; END_IF;
    #r := ("ROLL_State".M[32, 2] OR "ROLL_State".M[41, 3] OR "ROLL_State".M[41, 6] OR "ROLL_State".M[43, 2] OR "ROLL_State".M[44, 7] OR "ROLL_State".M[46, 2] OR "ROLL_State".M[47, 6] OR "ROLL_State".M[49, 2]);
    IF #r THEN "ROLL_State".M[41, 2] := FALSE; END_IF;
    // PB9, STEP 5 network 29
    #r := ((NOT "ROLL_State".M[110, 1]) AND (NOT "ROLL_State".M[110, 2]) AND "ROLL_State".M[35, 2] AND "ROLL_State".M[41, 2]);
    IF #r THEN "ROLL_State".M[41, 3] := TRUE; END_IF;
    #r := ("ROLL_State".M[32, 2] OR "ROLL_State".M[41, 4]);
    IF #r THEN "ROLL_State".M[41, 3] := FALSE; END_IF;
    // PB9, STEP 5 network 30
    #r := ("ROLL_IO".Input[13, 3] AND "ROLL_State".M[35, 2] AND "ROLL_State".M[41, 3] AND "ROLL_State".M[63, 1]);
    IF #r THEN "ROLL_State".M[41, 4] := TRUE; END_IF;
    #r := ("ROLL_State".M[32, 2] OR "ROLL_State".M[44, 7] OR "ROLL_State".M[50, 6] OR "ROLL_State".M[52, 0]);
    IF #r THEN "ROLL_State".M[41, 4] := FALSE; END_IF;
    // PB9, STEP 5 network 31
    #r := ((NOT "ROLL_IO".Input[11, 2]) AND (((NOT "ROLL_State".M[110, 0]) AND "ROLL_State".M[40, 1]) OR "ROLL_State".M[41, 2]) AND "ROLL_IO".Input[12, 5] AND "ROLL_IO".Input[12, 7] AND "ROLL_State".M[110, 1] AND "ROLL_State".M[35, 2]);
    IF #r THEN "ROLL_State".M[41, 6] := TRUE; END_IF;
    #r := ("ROLL_State".M[32, 2] OR "ROLL_State".M[41, 7]);
    IF #r THEN "ROLL_State".M[41, 6] := FALSE; END_IF;
    // PB9, STEP 5 network 32
    #r := ("ROLL_IO".Input[11, 2] AND "ROLL_IO".Input[11, 6] AND "ROLL_State".M[35, 2] AND "ROLL_State".M[41, 6]);
    IF #r THEN "ROLL_State".M[41, 7] := TRUE; END_IF;
    #r := ("ROLL_State".M[32, 2] OR "ROLL_State".M[42, 0]);
    IF #r THEN "ROLL_State".M[41, 7] := FALSE; END_IF;
    // PB9, STEP 5 network 33
    #r := ((NOT "ROLL_IO".Input[12, 1]) AND "ROLL_IO".Input[12, 5] AND "ROLL_State".M[35, 2] AND "ROLL_State".M[41, 7]);
    IF #r THEN "ROLL_State".M[42, 0] := TRUE; END_IF;
    #r := ("ROLL_State".M[32, 2] OR "ROLL_State".M[42, 1]);
    IF #r THEN "ROLL_State".M[42, 0] := FALSE; END_IF;
    // PB9, STEP 5 network 34
    #r := ("ROLL_IO".Input[12, 1] AND "ROLL_IO".Input[12, 7] AND "ROLL_State".M[35, 2] AND "ROLL_State".M[42, 0]);
    IF #r THEN "ROLL_State".M[42, 1] := TRUE; END_IF;
    #r := ("ROLL_State".M[32, 2] OR "ROLL_State".M[42, 2]);
    IF #r THEN "ROLL_State".M[42, 1] := FALSE; END_IF;
    // PB9, STEP 5 network 35
    #r := ("ROLL_State".M[35, 2] AND "ROLL_State".M[42, 1] AND "ROLL_State".S5Timers[1].Q);
    IF #r THEN "ROLL_State".M[42, 2] := TRUE; END_IF;
    #r := ("ROLL_State".M[32, 2] OR "ROLL_State".M[42, 3]);
    IF #r THEN "ROLL_State".M[42, 2] := FALSE; END_IF;
    // PB9, STEP 5 network 36
    #r := ("ROLL_State".M[35, 2] AND "ROLL_State".M[42, 2]);
    IF #r THEN "ROLL_State".M[42, 3] := TRUE; END_IF;
    #r := ("ROLL_State".M[32, 2] OR "ROLL_State".M[42, 4]);
    IF #r THEN "ROLL_State".M[42, 3] := FALSE; END_IF;
    // PB9, STEP 5 network 37
    #r := ((NOT "ROLL_IO".Input[12, 5]) AND (("ROLL_IO".Input[13, 3] AND "ROLL_State".M[63, 1]) OR (NOT "ROLL_State".M[111, 5])) AND "ROLL_State".M[35, 2] AND "ROLL_State".M[42, 3]);
    IF #r THEN "ROLL_State".M[42, 4] := TRUE; END_IF;
    #r := ("ROLL_State".M[32, 2] OR "ROLL_State".M[42, 5]);
    IF #r THEN "ROLL_State".M[42, 4] := FALSE; END_IF;
    // PB9, STEP 5 network 38
    #r := ("ROLL_IO".Input[12, 5] AND "ROLL_IO".Input[12, 7] AND "ROLL_State".M[35, 2] AND "ROLL_State".M[42, 4]);
    IF #r THEN "ROLL_State".M[42, 5] := TRUE; END_IF;
    #r := ("ROLL_State".M[32, 2] OR "ROLL_State".M[42, 6]);
    IF #r THEN "ROLL_State".M[42, 5] := FALSE; END_IF;
    // PB9, STEP 5 network 39
    #r := ("ROLL_State".M[35, 2] AND "ROLL_State".M[42, 5] AND "ROLL_State".S5Timers[2].Q);
    IF #r THEN "ROLL_State".M[42, 6] := TRUE; END_IF;
    #r := ("ROLL_State".M[32, 2] OR "ROLL_State".M[42, 7] OR "ROLL_State".M[43, 2] OR "ROLL_State".M[44, 7] OR "ROLL_State".M[46, 2] OR "ROLL_State".M[47, 6] OR "ROLL_State".M[49, 2]);
    IF #r THEN "ROLL_State".M[42, 6] := FALSE; END_IF;
    // PB9, STEP 5 network 40
    #r := ((NOT "ROLL_State".M[110, 2]) AND "ROLL_State".M[35, 2] AND "ROLL_State".M[42, 6]);
    IF #r THEN "ROLL_State".M[42, 7] := TRUE; END_IF;
    #r := ("ROLL_State".M[32, 2] OR "ROLL_State".M[43, 0]);
    IF #r THEN "ROLL_State".M[42, 7] := FALSE; END_IF;
    // PB9, STEP 5 network 41
    #r := ("ROLL_IO".Input[13, 3] AND "ROLL_State".M[35, 2] AND "ROLL_State".M[42, 7] AND "ROLL_State".M[63, 1]);
    IF #r THEN "ROLL_State".M[43, 0] := TRUE; END_IF;
    #r := ("ROLL_State".M[32, 2] OR "ROLL_State".M[44, 7] OR "ROLL_State".M[50, 6] OR "ROLL_State".M[52, 0]);
    IF #r THEN "ROLL_State".M[43, 0] := FALSE; END_IF;
    // PB9, STEP 5 network 42
    #r := ((NOT "ROLL_IO".Input[11, 3]) AND (((NOT "ROLL_State".M[110, 0]) AND (NOT "ROLL_State".M[110, 1]) AND "ROLL_State".M[40, 1]) OR ((NOT "ROLL_State".M[110, 1]) AND "ROLL_State".M[41, 2]) OR "ROLL_State".M[42, 6]) AND "ROLL_IO".Input[12, 5] AND "ROLL_IO".Input[12, 7] AND "ROLL_State".M[110, 2] AND "ROLL_State".M[35, 2]);
    IF #r THEN "ROLL_State".M[43, 2] := TRUE; END_IF;
    #r := ("ROLL_State".M[32, 2] OR "ROLL_State".M[43, 3]);
    IF #r THEN "ROLL_State".M[43, 2] := FALSE; END_IF;
    // PB9, STEP 5 network 43
    #r := ("ROLL_IO".Input[11, 3] AND "ROLL_IO".Input[11, 6] AND "ROLL_State".M[35, 2] AND "ROLL_State".M[43, 2]);
    IF #r THEN "ROLL_State".M[43, 3] := TRUE; END_IF;
    #r := ("ROLL_State".M[32, 2] OR "ROLL_State".M[43, 4]);
    IF #r THEN "ROLL_State".M[43, 3] := FALSE; END_IF;
    // PB9, STEP 5 network 44
    #r := ((NOT "ROLL_IO".Input[12, 1]) AND "ROLL_IO".Input[12, 5] AND "ROLL_State".M[35, 2] AND "ROLL_State".M[43, 3]);
    IF #r THEN "ROLL_State".M[43, 4] := TRUE; END_IF;
    #r := ("ROLL_State".M[32, 2] OR "ROLL_State".M[43, 5]);
    IF #r THEN "ROLL_State".M[43, 4] := FALSE; END_IF;
    // PB9, STEP 5 network 45
    #r := ("ROLL_IO".Input[12, 1] AND "ROLL_IO".Input[12, 7] AND "ROLL_State".M[35, 2] AND "ROLL_State".M[43, 4]);
    IF #r THEN "ROLL_State".M[43, 5] := TRUE; END_IF;
    #r := ("ROLL_State".M[32, 2] OR "ROLL_State".M[43, 6]);
    IF #r THEN "ROLL_State".M[43, 5] := FALSE; END_IF;
    // PB9, STEP 5 network 46
    #r := ("ROLL_State".M[35, 2] AND "ROLL_State".M[43, 5] AND "ROLL_State".S5Timers[1].Q);
    IF #r THEN "ROLL_State".M[43, 6] := TRUE; END_IF;
    #r := ("ROLL_State".M[32, 2] OR "ROLL_State".M[43, 7]);
    IF #r THEN "ROLL_State".M[43, 6] := FALSE; END_IF;
    // PB9, STEP 5 network 47
    #r := ("ROLL_State".M[35, 2] AND "ROLL_State".M[43, 6]);
    IF #r THEN "ROLL_State".M[43, 7] := TRUE; END_IF;
    #r := ("ROLL_State".M[32, 2] OR "ROLL_State".M[44, 0]);
    IF #r THEN "ROLL_State".M[43, 7] := FALSE; END_IF;
    // PB9, STEP 5 network 48
    #r := ((NOT "ROLL_IO".Input[12, 5]) AND (("ROLL_IO".Input[13, 3] AND "ROLL_State".M[63, 1]) OR (NOT "ROLL_State".M[111, 5])) AND "ROLL_State".M[35, 2] AND "ROLL_State".M[43, 7]);
    IF #r THEN "ROLL_State".M[44, 0] := TRUE; END_IF;
    #r := ("ROLL_State".M[32, 2] OR "ROLL_State".M[44, 1]);
    IF #r THEN "ROLL_State".M[44, 0] := FALSE; END_IF;
    // PB9, STEP 5 network 49
    #r := ("ROLL_IO".Input[12, 5] AND "ROLL_IO".Input[12, 7] AND "ROLL_State".M[35, 2] AND "ROLL_State".M[44, 0]);
    IF #r THEN "ROLL_State".M[44, 1] := TRUE; END_IF;
    #r := ("ROLL_State".M[32, 2] OR "ROLL_State".M[44, 2]);
    IF #r THEN "ROLL_State".M[44, 1] := FALSE; END_IF;
    // PB9, STEP 5 network 50
    #r := ("ROLL_State".M[35, 2] AND "ROLL_State".M[44, 1] AND "ROLL_State".S5Timers[2].Q);
    IF #r THEN "ROLL_State".M[44, 2] := TRUE; END_IF;
    #r := ("ROLL_State".M[32, 2] OR "ROLL_State".M[44, 3] OR "ROLL_State".M[44, 7] OR "ROLL_State".M[46, 2] OR "ROLL_State".M[47, 6] OR "ROLL_State".M[49, 2]);
    IF #r THEN "ROLL_State".M[44, 2] := FALSE; END_IF;
    // PB9, STEP 5 network 51
    #r := ("ROLL_State".M[35, 2] AND "ROLL_State".M[44, 2]);
    IF #r THEN "ROLL_State".M[44, 3] := TRUE; END_IF;
    #r := ("ROLL_State".M[32, 2] OR "ROLL_State".M[44, 4]);
    IF #r THEN "ROLL_State".M[44, 3] := FALSE; END_IF;
    // PB9, STEP 5 network 52
    #r := ("ROLL_IO".Input[13, 3] AND "ROLL_State".M[35, 2] AND "ROLL_State".M[44, 3] AND "ROLL_State".M[63, 1]);
    IF #r THEN "ROLL_State".M[44, 4] := TRUE; END_IF;
    #r := ("ROLL_State".M[32, 2] OR "ROLL_State".M[44, 7] OR "ROLL_State".M[50, 6] OR "ROLL_State".M[52, 0]);
    IF #r THEN "ROLL_State".M[44, 4] := FALSE; END_IF;
    // PB9, STEP 5 network 53
    #r := (((NOT "ROLL_State".M[110, 0]) AND (NOT "ROLL_State".M[110, 1]) AND (NOT "ROLL_State".M[110, 2]) AND "ROLL_State".M[40, 1]) OR ((NOT "ROLL_State".M[110, 1]) AND (NOT "ROLL_State".M[110, 2]) AND "ROLL_State".M[41, 4]) OR ((NOT "ROLL_State".M[110, 2]) AND "ROLL_State".M[43, 0]) OR "ROLL_State".M[44, 4]);
    "ROLL_State".M[240, 0] := #r;
    // PB9, STEP 5 network 54
    #r := ((NOT "ROLL_IO".Input[11, 4]) AND "ROLL_IO".Input[12, 5] AND "ROLL_IO".Input[12, 7] AND "ROLL_State".M[110, 3] AND "ROLL_State".M[240, 0] AND "ROLL_State".M[35, 2] AND "ROLL_State".M[63, 1]);
    IF #r THEN "ROLL_State".M[44, 7] := TRUE; END_IF;
    #r := ("ROLL_State".M[32, 2] OR "ROLL_State".M[45, 0]);
    IF #r THEN "ROLL_State".M[44, 7] := FALSE; END_IF;
    // PB9, STEP 5 network 55
    #r := ("ROLL_IO".Input[11, 4] AND "ROLL_IO".Input[11, 6] AND "ROLL_State".M[35, 2] AND "ROLL_State".M[44, 7]);
    IF #r THEN "ROLL_State".M[45, 0] := TRUE; END_IF;
    #r := ("ROLL_State".M[32, 2] OR "ROLL_State".M[45, 1]);
    IF #r THEN "ROLL_State".M[45, 0] := FALSE; END_IF;
    // PB9, STEP 5 network 56
    #r := ((NOT "ROLL_IO".Input[12, 1]) AND "ROLL_IO".Input[12, 5] AND "ROLL_State".M[35, 2] AND "ROLL_State".M[45, 0]);
    IF #r THEN "ROLL_State".M[45, 1] := TRUE; END_IF;
    #r := ("ROLL_State".M[32, 2] OR "ROLL_State".M[45, 2]);
    IF #r THEN "ROLL_State".M[45, 1] := FALSE; END_IF;
    // PB9, STEP 5 network 57
    #r := ("ROLL_IO".Input[12, 1] AND "ROLL_IO".Input[12, 7] AND "ROLL_State".M[35, 2] AND "ROLL_State".M[45, 1]);
    IF #r THEN "ROLL_State".M[45, 2] := TRUE; END_IF;
    #r := ("ROLL_State".M[32, 2] OR "ROLL_State".M[45, 3]);
    IF #r THEN "ROLL_State".M[45, 2] := FALSE; END_IF;
    // PB9, STEP 5 network 58
    #r := ("ROLL_State".M[35, 2] AND "ROLL_State".M[45, 2] AND "ROLL_State".S5Timers[1].Q);
    IF #r THEN "ROLL_State".M[45, 3] := TRUE; END_IF;
    #r := ("ROLL_State".M[32, 2] OR "ROLL_State".M[45, 4]);
    IF #r THEN "ROLL_State".M[45, 3] := FALSE; END_IF;
    // PB9, STEP 5 network 59
    #r := ("ROLL_State".M[35, 2] AND "ROLL_State".M[45, 3]);
    IF #r THEN "ROLL_State".M[45, 4] := TRUE; END_IF;
    #r := ("ROLL_State".M[32, 2] OR "ROLL_State".M[45, 5]);
    IF #r THEN "ROLL_State".M[45, 4] := FALSE; END_IF;
    // PB9, STEP 5 network 60
    #r := ((NOT "ROLL_IO".Input[12, 5]) AND "ROLL_State".M[35, 2] AND "ROLL_State".M[45, 4]);
    IF #r THEN "ROLL_State".M[45, 5] := TRUE; END_IF;
    #r := ("ROLL_State".M[32, 2] OR "ROLL_State".M[45, 6]);
    IF #r THEN "ROLL_State".M[45, 5] := FALSE; END_IF;
    // PB9, STEP 5 network 61
    #r := ("ROLL_IO".Input[12, 5] AND "ROLL_IO".Input[12, 7] AND "ROLL_State".M[35, 2] AND "ROLL_State".M[45, 5]);
    IF #r THEN "ROLL_State".M[45, 6] := TRUE; END_IF;
    #r := ("ROLL_State".M[32, 2] OR "ROLL_State".M[45, 7]);
    IF #r THEN "ROLL_State".M[45, 6] := FALSE; END_IF;
    // PB9, STEP 5 network 62
    #r := (("ROLL_State".M[0, 4] OR "ROLL_State".S5Timers[2].Q) AND "ROLL_State".M[35, 2] AND "ROLL_State".M[45, 6]);
    IF #r THEN "ROLL_State".M[45, 7] := TRUE; END_IF;
    #r := ("ROLL_State".M[32, 2] OR "ROLL_State".M[46, 0] OR "ROLL_State".M[46, 2] OR "ROLL_State".M[47, 6] OR "ROLL_State".M[49, 2]);
    IF #r THEN "ROLL_State".M[45, 7] := FALSE; END_IF;
    // PB9, STEP 5 network 63
    #r := ("ROLL_State".M[35, 2] AND "ROLL_State".M[45, 7]);
    IF #r THEN "ROLL_State".M[46, 0] := TRUE; END_IF;
    #r := ("ROLL_State".M[32, 2] OR "ROLL_State".M[46, 1]);
    IF #r THEN "ROLL_State".M[46, 0] := FALSE; END_IF;
    // PB9, STEP 5 network 64
    #r := ("ROLL_IO".Input[13, 3] AND "ROLL_State".M[35, 2] AND "ROLL_State".M[46, 0] AND "ROLL_State".M[63, 1]);
    IF #r THEN "ROLL_State".M[46, 1] := TRUE; END_IF;
    #r := ("ROLL_State".M[32, 2] OR "ROLL_State".M[50, 6] OR "ROLL_State".M[52, 0]);
    IF #r THEN "ROLL_State".M[46, 1] := FALSE; END_IF;
    // PB9, STEP 5 network 65
    RETURN;
END_FUNCTION

